(* IEC 61131-3 sources: brOscatLib/oscatBasic (part 6) *)

FUNCTION MIRROR : BOOL (* String *) (* http://www.oscat.de/images/OSCATBasic/oscat_basic333_en.pdf#page=174 *)
	VAR_INPUT
		STR : STRING[STRING_LENGTH];
	END_VAR
	VAR_IN_OUT
		RETVAL : STRING[STRING_LENGTH]; (*Return value of the function*)
	END_VAR
	VAR
		pi : REFERENCE TO ARRAY[1..255] OF BYTE;
		po : REFERENCE TO BYTE;
		lx : INT;
		i : INT;
	END_VAR
END_FUNCTION

FUNCTION MIX : REAL (* Signal processing *) (* http://www.oscat.de/images/OSCATBasic/oscat_basic333_en.pdf#page=281 *)
	VAR_INPUT
		A : REAL;
		B : REAL;
		M : REAL;
	END_VAR
END_FUNCTION

FUNCTION MODR : REAL (* Mathematical *) (* http://www.oscat.de/images/OSCATBasic/oscat_basic333_en.pdf#page=60 *)
	VAR_INPUT
		IN : REAL;
		DIVI : REAL;
	END_VAR
END_FUNCTION

FUNCTION MONTH_BEGIN : DATE (* Time and date *) (* http://www.oscat.de/images/OSCATBasic/oscat_basic333_en.pdf#page=129 *)
	VAR_INPUT
		IDATE : DATE;
	END_VAR
END_FUNCTION

FUNCTION MONTH_END : DATE (* Time and date *) (* http://www.oscat.de/images/OSCATBasic/oscat_basic333_en.pdf#page=130 *)
	VAR_INPUT
		IDATE : DATE;
	END_VAR
END_FUNCTION

FUNCTION MONTH_OF_DATE : INT (* Time and date *) (* http://www.oscat.de/images/OSCATBasic/oscat_basic333_en.pdf#page=130 *)
	VAR_INPUT
		IDATE : DATE;
	END_VAR
END_FUNCTION

FUNCTION MONTH_TO_STRING : BOOL (* String *) (* http://www.oscat.de/images/OSCATBasic/oscat_basic333_en.pdf#page=175 *)
	VAR_INPUT
		MTH : INT;
		LANG : INT;
		LX : INT;
	END_VAR
	VAR_IN_OUT
		RETVAL : STRING[10]; (*Return value of the function*)
	END_VAR
	VAR
		ly : INT;
	END_VAR
	VAR CONSTANT
		cMONTHS : ARRAY[1..3,1..12] OF STRING[10] := ['January','February','March','April','May','June','July','August','September','October','November','December','Januar','Februar','März','April','Mai','Juni','Juli','August','September','Oktober','November','Dezember','Janvier','Février','mars','Avril','Mai','Juin','Juillet','Août','Septembre','Octobre','Novembre','Decembre'];
		cMONTHS3 : ARRAY[1..3,1..12] OF STRING[3] := ['Jan','Feb','Mar','Apr','May','Jun','Jul','Aug','Sep','Oct','Nov','Dec','Jan','Feb','Mrz','Apr','Mai','Jun','Jul','Aug','Sep','Okt','Nov','Dez','Jan','Fev','Mar','Avr','Mai','Jun','Jul','Aou','Sep','Oct','Nov','Dec'];
	END_VAR
END_FUNCTION

FUNCTION MS_TO_BFT : INT (* Conversion *) (* http://www.oscat.de/images/OSCATBasic/oscat_basic333_en.pdf#page=368 *)
	VAR_INPUT
		MS : REAL;
	END_VAR
END_FUNCTION

FUNCTION MS_TO_KMH : REAL (* Conversion *) (* http://www.oscat.de/images/OSCATBasic/oscat_basic333_en.pdf#page=369 *)
	VAR_INPUT
		MS : REAL;
	END_VAR
END_FUNCTION

FUNCTION MULTIME : TIME (* Time and date *) (* http://www.oscat.de/images/OSCATBasic/oscat_basic333_en.pdf#page=130 *)
	VAR_INPUT
		T : TIME;
		M : REAL;
	END_VAR
END_FUNCTION

FUNCTION MULTI_IN : REAL (* Sensor *) (* http://www.oscat.de/images/OSCATBasic/oscat_basic333_en.pdf#page=317 *)
	VAR_INPUT
		IN_1 : REAL;
		IN_2 : REAL;
		IN_3 : REAL;
		DEFAULT : REAL;
		IN_MIN : REAL;
		IN_MAX : REAL;
		MODE : USINT;
	END_VAR
	VAR
		count : INT;
		F1 : BOOL;
		F2 : BOOL;
		F3 : BOOL;
	END_VAR
END_FUNCTION

FUNCTION MUL_ADD : REAL (* Mathematical *) (* http://www.oscat.de/images/OSCATBasic/oscat_basic333_en.pdf#page=61 *)
	VAR_INPUT
		X : REAL;
		K : REAL;
		O : REAL;
	END_VAR
END_FUNCTION

FUNCTION MUX_2 : BOOL (* Gate logic *) (* http://www.oscat.de/images/OSCATBasic/oscat_basic333_en.pdf#page=229 *)
	VAR_INPUT
		D0 : BOOL;
		D1 : BOOL;
		A0 : BOOL;
	END_VAR
END_FUNCTION

FUNCTION MUX_4 : BOOL (* Gate logic *) (* http://www.oscat.de/images/OSCATBasic/oscat_basic333_en.pdf#page=229 *)
	VAR_INPUT
		D0 : BOOL;
		D1 : BOOL;
		D2 : BOOL;
		D3 : BOOL;
		A0 : BOOL;
		A1 : BOOL;
	END_VAR
END_FUNCTION

FUNCTION MUX_R2 : REAL (* Signal processing *) (* http://www.oscat.de/images/OSCATBasic/oscat_basic333_en.pdf#page=281 *)
	VAR_INPUT
		IN0 : REAL;
		IN1 : REAL;
		A : BOOL;
	END_VAR
END_FUNCTION

FUNCTION MUX_R4 : REAL (* Signal processing *) (* http://www.oscat.de/images/OSCATBasic/oscat_basic333_en.pdf#page=282 *)
	VAR_INPUT
		IN0 : REAL;
		IN1 : REAL;
		IN2 : REAL;
		IN3 : REAL;
		A0 : BOOL;
		A1 : BOOL;
	END_VAR
END_FUNCTION

FUNCTION_BLOCK M_D (* Measurements *) (* http://www.oscat.de/images/OSCATBasic/oscat_basic333_en.pdf#page=341 *)
	VAR_INPUT
		START : BOOL;
		STOP : BOOL;
		TMAX : TIME := TIME#14400m0s0ms;
		RST : BOOL;
	END_VAR
	VAR_OUTPUT
		PT : TIME;
		ET : TIME;
		RUN : BOOL;
	END_VAR
	VAR
		edge_ : BOOL;
		T0 : TIME;
		tx : TIME;
		startup : BOOL;
	END_VAR
END_FUNCTION_BLOCK

FUNCTION_BLOCK M_T (* Measurements *) (* http://www.oscat.de/images/OSCATBasic/oscat_basic333_en.pdf#page=342 *)
	VAR_INPUT
		IN : BOOL;
		TMAX : TIME := TIME#14400m0s0ms;
		RST : BOOL;
	END_VAR
	VAR_OUTPUT
		PT : TIME;
		ET : TIME;
	END_VAR
	VAR
		edge_ : BOOL;
		start : TIME;
		tx : TIME;
	END_VAR
END_FUNCTION_BLOCK

FUNCTION_BLOCK M_TX (* Measurements *) (* http://www.oscat.de/images/OSCATBasic/oscat_basic333_en.pdf#page=342 *)
	VAR_INPUT
		IN : BOOL;
		TMAX : TIME := TIME#14400m0s0ms;
		RST : BOOL;
	END_VAR
	VAR_OUTPUT
		TH : TIME;
		TL : TIME;
		DC : REAL;
		F : REAL;
		ET : TIME;
	END_VAR
	VAR
		edge_ : BOOL;
		start : TIME;
		stop : TIME;
		tx : TIME;
		rise : BOOL;
		fall : BOOL;
		startup : BOOL;
	END_VAR
END_FUNCTION_BLOCK

FUNCTION NEGX : REAL (* Mathematical *) (* http://www.oscat.de/images/OSCATBasic/oscat_basic333_en.pdf#page=61 *)
	VAR_INPUT
		X : REAL;
	END_VAR
END_FUNCTION

FUNCTION OCT_TO_BYTE : BYTE (* String *) (* http://www.oscat.de/images/OSCATBasic/oscat_basic333_en.pdf#page=175 *)
	VAR_INPUT
		OCT : STRING[10];
	END_VAR
	VAR
		pt : REFERENCE TO BYTE;
		i : INT;
		X : BYTE;
		stop : INT;
		intX : USINT;
	END_VAR
END_FUNCTION

FUNCTION OCT_TO_DWORD : DWORD (* String *) (* http://www.oscat.de/images/OSCATBasic/oscat_basic333_en.pdf#page=176 *)
	VAR_INPUT
		OCT : STRING[20];
	END_VAR
	VAR
		pt : REFERENCE TO BYTE;
		i : INT;
		X : BYTE;
		stop : INT;
		intX : USINT;
		temp : UDINT;
	END_VAR
END_FUNCTION

FUNCTION OFFSET : REAL (* Signal processing *) (* http://www.oscat.de/images/OSCATBasic/oscat_basic333_en.pdf#page=282 *)
	VAR_INPUT
		X : REAL;
		O1 : BOOL;
		O2 : BOOL;
		O3 : BOOL;
		O4 : BOOL;
		D : BOOL;
		OFFSET_1 : REAL;
		OFFSET_2 : REAL;
		OFFSET_3 : REAL;
		OFFSET_4 : REAL;
		DEFAULT : REAL;
	END_VAR
END_FUNCTION

FUNCTION OFFSET2 : REAL (* Signal processing *) (* http://www.oscat.de/images/OSCATBasic/oscat_basic333_en.pdf#page=285 *)
	VAR_INPUT
		X : REAL;
		O1 : BOOL;
		O2 : BOOL;
		O3 : BOOL;
		O4 : BOOL;
		D : BOOL;
		OFFSET_1 : REAL;
		OFFSET_2 : REAL;
		OFFSET_3 : REAL;
		OFFSET_4 : REAL;
		DEFAULT : REAL;
	END_VAR
END_FUNCTION

FUNCTION OM_TO_F : REAL (* Conversion *) (* http://www.oscat.de/images/OSCATBasic/oscat_basic333_en.pdf#page=369 *)
	VAR_INPUT
		OM : REAL;
	END_VAR
END_FUNCTION

FUNCTION_BLOCK ONTIME (* Measurements *) (* http://www.oscat.de/images/OSCATBasic/oscat_basic333_en.pdf#page=346 *)
	VAR_INPUT
		IN : BOOL;
		RST : BOOL;
	END_VAR
	VAR_IN_OUT
		SECONDS : UDINT;
		CYCLES : UDINT;
	END_VAR
	VAR
		tx : UDINT;
		last : UDINT;
		edge_ : BOOL;
		init : BOOL;
		ms : UDINT;
	END_VAR
END_FUNCTION_BLOCK

FUNCTION OSCAT_VERSION : DWORD (* Other *) (* http://www.oscat.de/images/OSCATBasic/oscat_basic333_en.pdf#page=37 *)
	VAR_INPUT
		IN : BOOL;
	END_VAR
END_FUNCTION

FUNCTION OVERRIDE : REAL (* Signal processing *) (* http://www.oscat.de/images/OSCATBasic/oscat_basic333_en.pdf#page=286 *)
	VAR_INPUT
		X1 : REAL;
		X2 : REAL;
		X3 : REAL;
		E1 : BOOL;
		E2 : BOOL;
		E3 : BOOL;
	END_VAR
END_FUNCTION

FUNCTION PARITY : BOOL (* Gate logic *) (* http://www.oscat.de/images/OSCATBasic/oscat_basic333_en.pdf#page=230 *)
	VAR_INPUT
		IN : DWORD;
	END_VAR
END_FUNCTION

FUNCTION_BLOCK PARSET (* Automation *) (* http://www.oscat.de/images/OSCATBasic/oscat_basic333_en.pdf#page=466 *)
	VAR_INPUT
		A0 : BOOL;
		A1 : BOOL;
		X01 : REAL;
		X02 : REAL;
		X03 : REAL;
		X04 : REAL;
		X11 : REAL;
		X12 : REAL;
		X13 : REAL;
		X14 : REAL;
		X21 : REAL;
		X22 : REAL;
		X23 : REAL;
		X24 : REAL;
		X31 : REAL;
		X32 : REAL;
		X33 : REAL;
		X34 : REAL;
		TC : TIME;
	END_VAR
	VAR_OUTPUT
		P1 : REAL;
		P2 : REAL;
		P3 : REAL;
		P4 : REAL;
	END_VAR
	VAR
		X : ARRAY[0..3,1..4] OF REAL;
		S1 : REAL;
		S2 : REAL;
		S3 : REAL;
		S4 : REAL;
		tx : UDINT;
		last : UDINT;
		start : BOOL;
		set : USINT;
		init : BOOL;
	END_VAR
END_FUNCTION_BLOCK

FUNCTION_BLOCK PARSET2 (* Automation *) (* http://www.oscat.de/images/OSCATBasic/oscat_basic333_en.pdf#page=467 *)
	VAR_INPUT
		X : REAL;
		X01 : REAL;
		X02 : REAL;
		X03 : REAL;
		X04 : REAL;
		X11 : REAL;
		X12 : REAL;
		X13 : REAL;
		X14 : REAL;
		X21 : REAL;
		X22 : REAL;
		X23 : REAL;
		X24 : REAL;
		X31 : REAL;
		X32 : REAL;
		X33 : REAL;
		X34 : REAL;
		L1 : REAL;
		L2 : REAL;
		L3 : REAL;
		TC : TIME;
	END_VAR
	VAR_OUTPUT
		P1 : REAL;
		P2 : REAL;
		P3 : REAL;
		P4 : REAL;
	END_VAR
	VAR
		Pset : PARSET;
		init : BOOL;
	END_VAR
END_FUNCTION_BLOCK

FUNCTION PERIOD : BOOL (* Time and date *) (* http://www.oscat.de/images/OSCATBasic/oscat_basic333_en.pdf#page=131 *)
	VAR_INPUT
		D1 : DATE;
		DX : DATE;
		D2 : DATE;
	END_VAR
	VAR
		day1 : INT;
		day2 : INT;
		dayx : INT;
	END_VAR
END_FUNCTION

FUNCTION PERIOD2 : BOOL (* Time and date *) (* http://www.oscat.de/images/OSCATBasic/oscat_basic333_en.pdf#page=131 *)
	VAR_INPUT
		DP : ARRAY[0..3,0..1] OF DATE;
		DX : DATE;
	END_VAR
END_FUNCTION

FUNCTION_BLOCK PIN_CODE (* Others *) (* http://www.oscat.de/images/OSCATBasic/oscat_basic333_en.pdf#page=231 *)
	VAR_INPUT
		CB : BYTE;
		E : BOOL;
		PIN : STRING[8];
	END_VAR
	VAR_OUTPUT
		TP : BOOL;
	END_VAR
	VAR
		POS : INT := 1;
	END_VAR
END_FUNCTION_BLOCK

FUNCTION POLYNOM_INT : REAL (* Functions *) (* http://www.oscat.de/images/OSCATBasic/oscat_basic333_en.pdf#page=102 *)
	VAR_INPUT
		X : REAL;
		XY : ARRAY[1..5,0..1] OF REAL;
		PTS : INT;
	END_VAR
	VAR
		I : INT;
		J : INT;
		stop : INT;
	END_VAR
END_FUNCTION

FUNCTION_BLOCK PRESSURE (* Conversion *) (* http://www.oscat.de/images/OSCATBasic/oscat_basic333_en.pdf#page=371 *)
	VAR_INPUT
		MWS : REAL;
		TORR : REAL;
		ATT : REAL;
		ATM : REAL;
		PA : REAL;
		BAR : REAL;
	END_VAR
	VAR_OUTPUT
		YMWS : REAL;
		YTORR : REAL;
		YATT : REAL;
		YATM : REAL;
		YPA : REAL;
		YBAR : REAL;
	END_VAR
END_FUNCTION_BLOCK

FUNCTION PT_TO_F : REAL (* Conversion *) (* http://www.oscat.de/images/OSCATBasic/oscat_basic333_en.pdf#page=372 *)
	VAR_INPUT
		PT : TIME;
	END_VAR
END_FUNCTION

FUNCTION_BLOCK PWM_DC (* Signal generators *) (* http://www.oscat.de/images/OSCATBasic/oscat_basic333_en.pdf#page=263 *)
	VAR_INPUT
		F : REAL;
		DC : REAL;
	END_VAR
	VAR_OUTPUT
		Q : BOOL;
	END_VAR
	VAR
		clk : CLK_PRG;
		pulse : TP_X;
		tmp : REAL;
	END_VAR
END_FUNCTION_BLOCK

FUNCTION_BLOCK PWM_PW (* Signal generators *) (* http://www.oscat.de/images/OSCATBasic/oscat_basic333_en.pdf#page=264 *)
	VAR_INPUT
		F : REAL;
		PW : TIME;
	END_VAR
	VAR_OUTPUT
		Q : BOOL;
	END_VAR
	VAR
		clk : CLK_PRG;
		pulse : TP_X;
	END_VAR
END_FUNCTION_BLOCK

FUNCTION R2_ABS : BOOL (* Double Precision *) (* http://www.oscat.de/images/OSCATBasic/oscat_basic333_en.pdf#page=93 *)
	VAR_INPUT
		X : REAL2;
	END_VAR
	VAR_IN_OUT
		RETVAL : REAL2; (*Return value of the function*)
	END_VAR
END_FUNCTION

FUNCTION R2_ADD : BOOL (* Double Precision *) (* http://www.oscat.de/images/OSCATBasic/oscat_basic333_en.pdf#page=93 *)
	VAR_INPUT
		X : REAL2;
		Y : REAL;
	END_VAR
	VAR_IN_OUT
		RETVAL : REAL2; (*Return value of the function*)
	END_VAR
	VAR
		temp : REAL;
	END_VAR
END_FUNCTION

FUNCTION R2_ADD2 : BOOL (* Double Precision *) (* http://www.oscat.de/images/OSCATBasic/oscat_basic333_en.pdf#page=94 *)
	VAR_INPUT
		X : REAL2;
		Y : REAL2;
	END_VAR
	VAR_IN_OUT
		RETVAL : REAL2; (*Return value of the function*)
	END_VAR
END_FUNCTION

FUNCTION R2_MUL : BOOL (* Double Precision *) (* http://www.oscat.de/images/OSCATBasic/oscat_basic333_en.pdf#page=94 *)
	VAR_INPUT
		X : REAL2;
		Y : REAL;
	END_VAR
	VAR_IN_OUT
		RETVAL : REAL2; (*Return value of the function*)
	END_VAR
END_FUNCTION

FUNCTION R2_SET : BOOL (* Double Precision *) (* http://www.oscat.de/images/OSCATBasic/oscat_basic333_en.pdf#page=95 *)
	VAR_INPUT
		X : REAL;
	END_VAR
	VAR_IN_OUT
		RETVAL : REAL2; (*Return value of the function*)
	END_VAR
END_FUNCTION

FUNCTION RAD : REAL (* Mathematical *) (* http://www.oscat.de/images/OSCATBasic/oscat_basic333_en.pdf#page=61 *)
	VAR_INPUT
		DEG : REAL;
	END_VAR
END_FUNCTION

FUNCTION RANGE_TO_BYTE : BYTE (* Signal processing *) (* http://www.oscat.de/images/OSCATBasic/oscat_basic333_en.pdf#page=288 *)
	VAR_INPUT
		X : REAL;
		LOW : REAL;
		HIGH : REAL;
	END_VAR
END_FUNCTION

FUNCTION RANGE_TO_WORD : WORD (* Signal processing *) (* http://www.oscat.de/images/OSCATBasic/oscat_basic333_en.pdf#page=288 *)
	VAR_INPUT
		X : REAL;
		LOW : REAL;
		HIGH : REAL;
	END_VAR
END_FUNCTION

FUNCTION RDM : REAL (* Mathematical *) (* http://www.oscat.de/images/OSCATBasic/oscat_basic333_en.pdf#page=62 *)
	VAR_INPUT
		LAST : REAL;
	END_VAR
	VAR
		tn : UDINT;
		tc : INT;
	END_VAR
END_FUNCTION

FUNCTION RDM2 : INT (* Mathematical *) (* http://www.oscat.de/images/OSCATBasic/oscat_basic333_en.pdf#page=62 *)
	VAR_INPUT
		LAST : INT;
		LOW : INT;
		HIGH : INT;
	END_VAR
END_FUNCTION

FUNCTION RDMDW : DWORD (* Mathematical *) (* http://www.oscat.de/images/OSCATBasic/oscat_basic333_en.pdf#page=63 *)
	VAR_INPUT
		LAST : DWORD;
	END_VAR
	VAR
		RX : REAL;
		M : REAL;
	END_VAR
END_FUNCTION

FUNCTION REAL_TO_DW : DWORD (* Gate logic *) (* http://www.oscat.de/images/OSCATBasic/oscat_basic333_en.pdf#page=231 *)
	VAR_INPUT
		X : REAL;
	END_VAR
	VAR
		pt : REFERENCE TO DWORD;
	END_VAR
END_FUNCTION

FUNCTION REAL_TO_FRAC : BOOL (* Mathematical *) (* http://www.oscat.de/images/OSCATBasic/oscat_basic333_en.pdf#page=64 *)
	VAR_INPUT
		X : REAL; (* in einen Bruch umzuwandelnder Wert *)
		N : INT; (* maximale Größe des Nenners *)
	END_VAR
	VAR_IN_OUT
		RETVAL : FRACTION; (*Return value of the function*)
	END_VAR
	VAR
		temp : DINT; (* Merker für Berechnungen *)
		sign : BOOL; (* Vorzeichen vom Eingangswert *)
		X_gerundet : DINT; (* Wert von Bruch, auf ganze Zahl gerundet *)
		X_ohne_Nachkomma : REAL; (* Wert von Bruch, ohne Nachkommastellen *)
		Numerator : DINT := 1; (* Initialwert Zaehler  *)
		Denominator : DINT := 0; (* Initialwert Nenner *)
		Numerator_old : DINT := 0; (* Initialwert Zaehler der letzten Berechnung  *)
		Denominator_old : DINT := 1; (* Initialwert Zaehler der letzten Berechnung   *)
	END_VAR
END_FUNCTION

FUNCTION REAL_TO_STRF : BOOL (* String *) (* http://www.oscat.de/images/OSCATBasic/oscat_basic333_en.pdf#page=176 *)
	VAR_INPUT
		IN : REAL;
		N : INT;
		D : STRING[1];
	END_VAR
	VAR_IN_OUT
		RETVAL : STRING[20]; (*Return value of the function*)
	END_VAR
	VAR
		O : REAL;
		i : INT;
	END_VAR
END_FUNCTION

FUNCTION REFLECT : DWORD (* Gate logic *) (* http://www.oscat.de/images/OSCATBasic/oscat_basic333_en.pdf#page=232 *)
	VAR_INPUT
		D : DWORD;
		L : INT;
	END_VAR
	VAR
		i : INT;
	END_VAR
END_FUNCTION

FUNCTION REFRACTION : REAL (* Time and date *) (* http://www.oscat.de/images/OSCATBasic/oscat_basic333_en.pdf#page=132 *)
	VAR_INPUT
		ELEV : REAL;
	END_VAR
END_FUNCTION

FUNCTION REPLACE_ALL : BOOL (* String *) (* http://www.oscat.de/images/OSCATBasic/oscat_basic333_en.pdf#page=177 *)
	VAR_INPUT
		STR : STRING[STRING_LENGTH];
		SRC : STRING[STRING_LENGTH];
		REP : STRING[STRING_LENGTH];
	END_VAR
	VAR_IN_OUT
		RETVAL : STRING[STRING_LENGTH]; (*Return value of the function*)
	END_VAR
	VAR
		pos : INT;
		lp : INT;
		lx : INT;
	END_VAR
END_FUNCTION

FUNCTION REPLACE_CHARS : BOOL (* String *) (* http://www.oscat.de/images/OSCATBasic/oscat_basic333_en.pdf#page=177 *)
	VAR_INPUT
		STR : STRING[STRING_LENGTH];
		SRC : STRING[255];
		REP : STRING[255];
	END_VAR
	VAR_IN_OUT
		RETVAL : STRING[STRING_LENGTH]; (*Return value of the function*)
	END_VAR
	VAR
		a : INT;
		b : INT;
		c : STRING[1];
		stp : INT;
	END_VAR
END_FUNCTION

FUNCTION REPLACE_UML : BOOL (* String *) (* http://www.oscat.de/images/OSCATBasic/oscat_basic333_en.pdf#page=178 *)
	VAR_INPUT
		STR : STRING[STRING_LENGTH];
	END_VAR
	VAR_IN_OUT
		RETVAL : STRING[STRING_LENGTH]; (*Return value of the function*)
	END_VAR
	VAR
		L : INT;
		pt : REFERENCE TO BYTE;
		pto : REFERENCE TO BYTE;
		ptm : REFERENCE TO BYTE;
		pt1 : REFERENCE TO BYTE;
		pt2 : REFERENCE TO BYTE;
		su : STRING[2];
		pos : INT;
	END_VAR
END_FUNCTION

FUNCTION RES_NI : REAL (* Sensor *) (* http://www.oscat.de/images/OSCATBasic/oscat_basic333_en.pdf#page=318 *)
	VAR_INPUT
		T : REAL;
		R0 : REAL;
	END_VAR
	VAR CONSTANT
		A : REAL := 0.5485;
		B : REAL := 0.000665;
		C : REAL := 2.805E-09;
	END_VAR
	VAR
		T2 : REAL;
	END_VAR
END_FUNCTION

FUNCTION RES_NTC : REAL (* Sensor *) (* http://www.oscat.de/images/OSCATBasic/oscat_basic333_en.pdf#page=319 *)
	VAR_INPUT
		T : REAL;
		RN : REAL;
		B : REAL;
	END_VAR
END_FUNCTION

FUNCTION RES_PT : REAL (* Sensor *) (* http://www.oscat.de/images/OSCATBasic/oscat_basic333_en.pdf#page=322 *)
	VAR_INPUT
		T : REAL;
		R0 : REAL;
	END_VAR
	VAR CONSTANT
		A : REAL := 0.00390802;
		B : REAL := -5.802E-07;
		C : REAL := -4.2735E-12;
	END_VAR
	VAR
		T2 : REAL;
	END_VAR
END_FUNCTION

FUNCTION RES_SI : REAL (* Sensor *) (* http://www.oscat.de/images/OSCATBasic/oscat_basic333_en.pdf#page=323 *)
	VAR_INPUT
		T : REAL;
		RS : REAL;
		TS : REAL;
	END_VAR
	VAR CONSTANT
		A : REAL := 0.00764;
		B : REAL := 1.66E-05;
	END_VAR
	VAR
		TX : REAL;
	END_VAR
END_FUNCTION

FUNCTION REVERSE : BYTE (* Gate logic *) (* http://www.oscat.de/images/OSCATBasic/oscat_basic333_en.pdf#page=232 *)
	VAR_INPUT
		IN : BYTE;
	END_VAR
END_FUNCTION

FUNCTION_BLOCK RMP_B (* Signal generators *) (* http://www.oscat.de/images/OSCATBasic/oscat_basic333_en.pdf#page=264 *)
	VAR_INPUT
		SET : BOOL;
		PT : TIME;
		E : BOOL := TRUE;
		UP : BOOL := TRUE;
		RST : BOOL;
	END_VAR
	VAR_OUTPUT
		OUT : BYTE;
		BUSY : BOOL;
		HIGH : BOOL;
		LOW : BOOL;
	END_VAR
	VAR
		rmp : _RMP_B;
	END_VAR
END_FUNCTION_BLOCK

FUNCTION_BLOCK RMP_SOFT (* Signal generators *) (* http://www.oscat.de/images/OSCATBasic/oscat_basic333_en.pdf#page=266 *)
	VAR_INPUT
		IN : BOOL;
		VAL : BYTE;
		PT_ON : TIME;
		PT_OFF : TIME;
	END_VAR
	VAR_OUTPUT
		OUT : BYTE;
	END_VAR
	VAR
		rmp : _RMP_B;
		tmp : BYTE;
	END_VAR
END_FUNCTION_BLOCK

FUNCTION_BLOCK RMP_W (* Signal generators *) (* http://www.oscat.de/images/OSCATBasic/oscat_basic333_en.pdf#page=267 *)
	VAR_INPUT
		SET : BOOL;
		PT : TIME;
		E : BOOL := TRUE;
		UP : BOOL := TRUE;
		RST : BOOL;
	END_VAR
	VAR_OUTPUT
		OUT : WORD;
		BUSY : BOOL;
		HIGH : BOOL;
		LOW : BOOL;
	END_VAR
	VAR
		rmp : _RMP_W;
	END_VAR
END_FUNCTION_BLOCK

FUNCTION RND : REAL (* Mathematical *) (* http://www.oscat.de/images/OSCATBasic/oscat_basic333_en.pdf#page=64 *)
	VAR_INPUT
		X : REAL;
		N : INT;
	END_VAR
	VAR
		M : REAL;
	END_VAR
END_FUNCTION

FUNCTION ROUND : REAL (* Mathematical *) (* http://www.oscat.de/images/OSCATBasic/oscat_basic333_en.pdf#page=65 *)
	VAR_INPUT
		IN : REAL;
		N : INT;
	END_VAR
	VAR
		X : REAL;
	END_VAR
	VAR CONSTANT
		cDECADES : ARRAY[0..8] OF REAL := [1,10,100,1000,10000,100000,1000000,10000000,100000000];
	END_VAR
END_FUNCTION

FUNCTION_BLOCK RTC_2 (* Time and date *) (* http://www.oscat.de/images/OSCATBasic/oscat_basic333_en.pdf#page=133 *)
	VAR_INPUT
		SET : BOOL;
		SDT : DATE_AND_TIME;
		SMS : INT;
		DEN : BOOL;
		OFS : INT;
	END_VAR
	VAR_OUTPUT
		UDT : DATE_AND_TIME;
		LOCAL_DT : DATE_AND_TIME;
		DSO : BOOL;
		XMS : INT;
	END_VAR
	VAR
		RT : RTC_MS;
	END_VAR
END_FUNCTION_BLOCK

FUNCTION_BLOCK RTC_MS (* Time and date *) (* http://www.oscat.de/images/OSCATBasic/oscat_basic333_en.pdf#page=134 *)
	VAR_INPUT
		SET : BOOL;
		SDT : DATE_AND_TIME;
		SMS : INT;
	END_VAR
	VAR_OUTPUT
		XDT : DATE_AND_TIME;
		XMS : INT;
	END_VAR
	VAR
		init : BOOL;
		last : UDINT;
		Tx : UDINT;
	END_VAR
END_FUNCTION_BLOCK

FUNCTION SCALE : REAL (* Signal processing *) (* http://www.oscat.de/images/OSCATBasic/oscat_basic333_en.pdf#page=288 *)
	VAR_INPUT
		X : REAL;
		K : REAL;
		O : REAL;
		MX : REAL;
		MN : REAL;
	END_VAR
END_FUNCTION

FUNCTION SCALE_B : REAL (* Signal processing *) (* http://www.oscat.de/images/OSCATBasic/oscat_basic333_en.pdf#page=289 *)
	VAR_INPUT
		X : BYTE;
		I_LO : BYTE;
		I_HI : BYTE;
		O_LO : REAL;
		O_HI : REAL;
	END_VAR
	VAR
		_I_HI : USINT;
		_I_LO : USINT;
	END_VAR
END_FUNCTION

FUNCTION SCALE_B2 : REAL (* Signal processing *) (* http://www.oscat.de/images/OSCATBasic/oscat_basic333_en.pdf#page=290 *)
	VAR_INPUT
		IN1 : BYTE;
		IN2 : BYTE;
		K : REAL;
		O : REAL;
		IN1_MIN : REAL;
		IN1_MAX : REAL := 1000;
		IN2_MIN : REAL;
		IN2_MAX : REAL := 1000;
	END_VAR
END_FUNCTION

FUNCTION SCALE_B4 : REAL (* Signal processing *) (* http://www.oscat.de/images/OSCATBasic/oscat_basic333_en.pdf#page=291 *)
	VAR_INPUT
		IN1 : BYTE;
		IN2 : BYTE;
		IN3 : BYTE;
		IN4 : BYTE;
		K : REAL;
		O : REAL;
		IN1_MIN : REAL;
		IN1_MAX : REAL := 1000;
		IN2_MIN : REAL;
		IN2_MAX : REAL := 1000;
		IN3_MIN : REAL;
		IN3_MAX : REAL := 1000;
		IN4_MIN : REAL;
		IN4_MAX : REAL := 1000;
	END_VAR
END_FUNCTION

FUNCTION SCALE_B8 : REAL (* Signal processing *) (* http://www.oscat.de/images/OSCATBasic/oscat_basic333_en.pdf#page=292 *)
	VAR_INPUT
		IN1 : BYTE;
		IN2 : BYTE;
		IN3 : BYTE;
		IN4 : BYTE;
		IN5 : BYTE;
		IN6 : BYTE;
		IN7 : BYTE;
		IN8 : BYTE;
		K : REAL;
		O : REAL;
		IN1_MIN : REAL;
		IN1_MAX : REAL := 1000;
		IN2_MIN : REAL;
		IN2_MAX : REAL := 1000;
		IN3_MIN : REAL;
		IN3_MAX : REAL := 1000;
		IN4_MIN : REAL;
		IN4_MAX : REAL := 1000;
		IN5_MIN : REAL;
		IN5_MAX : REAL := 1000;
		IN6_MIN : REAL;
		IN6_MAX : REAL := 1000;
		IN7_MIN : REAL;
		IN7_MAX : REAL := 1000;
		IN8_MIN : REAL;
		IN8_MAX : REAL := 1000;
	END_VAR
END_FUNCTION

FUNCTION SCALE_D : REAL (* Signal processing *) (* http://www.oscat.de/images/OSCATBasic/oscat_basic333_en.pdf#page=293 *)
	VAR_INPUT
		X : DWORD;
		I_LO : DWORD;
		I_HI : DWORD;
		O_LO : REAL;
		O_HI : REAL;
	END_VAR
	VAR
		_I_HI : UDINT;
		_I_LO : UDINT;
	END_VAR
END_FUNCTION

FUNCTION SCALE_R : REAL (* Signal processing *) (* http://www.oscat.de/images/OSCATBasic/oscat_basic333_en.pdf#page=294 *)
	VAR_INPUT
		X : REAL;
		I_LO : REAL;
		I_HI : REAL;
		O_LO : REAL;
		O_HI : REAL;
	END_VAR
END_FUNCTION

FUNCTION SCALE_X2 : REAL (* Signal processing *) (* http://www.oscat.de/images/OSCATBasic/oscat_basic333_en.pdf#page=295 *)
	VAR_INPUT
		IN1 : BOOL;
		IN2 : BOOL;
		K : REAL;
		O : REAL;
		IN1_MIN : REAL;
		IN1_MAX : REAL := 1000;
		IN2_MIN : REAL;
		IN2_MAX : REAL := 1000;
	END_VAR
END_FUNCTION

FUNCTION SCALE_X4 : REAL (* Signal processing *) (* http://www.oscat.de/images/OSCATBasic/oscat_basic333_en.pdf#page=296 *)
	VAR_INPUT
		IN1 : BOOL;
		IN2 : BOOL;
		IN3 : BOOL;
		IN4 : BOOL;
		K : REAL;
		O : REAL;
		IN1_MIN : REAL;
		IN1_MAX : REAL := 1000;
		IN2_MIN : REAL;
		IN2_MAX : REAL := 1000;
		IN3_MIN : REAL;
		IN3_MAX : REAL := 1000;
		IN4_MIN : REAL;
		IN4_MAX : REAL := 1000;
	END_VAR
END_FUNCTION

FUNCTION SCALE_X8 : REAL (* Signal processing *) (* http://www.oscat.de/images/OSCATBasic/oscat_basic333_en.pdf#page=297 *)
	VAR_INPUT
		IN1 : BOOL;
		IN2 : BOOL;
		IN3 : BOOL;
		IN4 : BOOL;
		IN5 : BOOL;
		IN6 : BOOL;
		IN7 : BOOL;
		IN8 : BOOL;
		K : REAL;
		O : REAL;
		IN1_MIN : REAL;
		IN1_MAX : REAL := 1000;
		IN2_MIN : REAL;
		IN2_MAX : REAL := 1000;
		IN3_MIN : REAL;
		IN3_MAX : REAL := 1000;
		IN4_MIN : REAL;
		IN4_MAX : REAL := 1000;
		IN5_MIN : REAL;
		IN5_MAX : REAL := 1000;
		IN6_MIN : REAL;
		IN6_MAX : REAL := 1000;
		IN7_MIN : REAL;
		IN7_MAX : REAL := 1000;
		IN8_MIN : REAL;
		IN8_MAX : REAL := 1000;
	END_VAR
END_FUNCTION

FUNCTION_BLOCK SCHEDULER (* Generators *) (* http://www.oscat.de/images/OSCATBasic/oscat_basic333_en.pdf#page=198 *)
	VAR_INPUT
		E0 : BOOL;
		E1 : BOOL;
		E2 : BOOL;
		E3 : BOOL;
		T0 : TIME;
		T1 : TIME;
		T2 : TIME;
		T3 : TIME;
	END_VAR
	VAR_OUTPUT
		Q0 : BOOL;
		Q1 : BOOL;
		Q2 : BOOL;
		Q3 : BOOL;
	END_VAR
	VAR
		init : BOOL;
		s0 : TIME;
		s1 : TIME;
		s2 : TIME;
		s3 : TIME;
		tx : TIME;
		c : INT;
	END_VAR
END_FUNCTION_BLOCK

FUNCTION_BLOCK SCHEDULER_2 (* Generators *) (* http://www.oscat.de/images/OSCATBasic/oscat_basic333_en.pdf#page=198 *)
	VAR_INPUT
		E0 : BOOL;
		E1 : BOOL;
		E2 : BOOL;
		E3 : BOOL;
		C0 : UINT;
		C1 : UINT;
		C2 : UINT;
		C3 : UINT;
		O0 : UINT;
		O1 : UINT;
		O2 : UINT;
		O3 : UINT;
	END_VAR
	VAR_OUTPUT
		Q0 : BOOL;
		Q1 : BOOL;
		Q2 : BOOL;
		Q3 : BOOL;
	END_VAR
	VAR
		sx : UINT;
	END_VAR
END_FUNCTION_BLOCK

FUNCTION SDT_TO_DATE : DATE (* Time and date *) (* http://www.oscat.de/images/OSCATBasic/oscat_basic333_en.pdf#page=134 *)
	VAR_INPUT
		DTI : SDT;
	END_VAR
END_FUNCTION

FUNCTION SDT_TO_DT : DATE_AND_TIME (* Time and date *) (* http://www.oscat.de/images/OSCATBasic/oscat_basic333_en.pdf#page=135 *)
	VAR_INPUT
		DTI : SDT;
	END_VAR
END_FUNCTION

FUNCTION SDT_TO_TOD : TIME_OF_DAY (* Time and date *) (* http://www.oscat.de/images/OSCATBasic/oscat_basic333_en.pdf#page=135 *)
	VAR_INPUT
		DTI : SDT;
	END_VAR
END_FUNCTION

FUNCTION SECOND : REAL (* Time and date *) (* http://www.oscat.de/images/OSCATBasic/oscat_basic333_en.pdf#page=135 *)
	VAR_INPUT
		ITOD : TIME_OF_DAY;
	END_VAR
END_FUNCTION

FUNCTION SECOND_OF_DT : INT (* Time and date *) (* http://www.oscat.de/images/OSCATBasic/oscat_basic333_en.pdf#page=136 *)
	VAR_INPUT
		XDT : DATE_AND_TIME;
	END_VAR
END_FUNCTION

FUNCTION SECOND_TO_TIME : TIME (* Time and date *) (* http://www.oscat.de/images/OSCATBasic/oscat_basic333_en.pdf#page=136 *)
	VAR_INPUT
		IN : REAL;
	END_VAR
END_FUNCTION

FUNCTION_BLOCK SEL2_OF_3 (* Signal processing *) (* http://www.oscat.de/images/OSCATBasic/oscat_basic333_en.pdf#page=298 *)
	VAR_INPUT
		IN1 : REAL;
		IN2 : REAL;
		IN3 : REAL;
		D : REAL;
	END_VAR
	VAR_OUTPUT
		Y : REAL;
		W : INT;
		E : BOOL;
	END_VAR
	VAR
		D12 : BOOL;
		D23 : BOOL;
		D31 : BOOL;
	END_VAR
END_FUNCTION_BLOCK

FUNCTION_BLOCK SEL2_OF_3B (* Signal processing *) (* http://www.oscat.de/images/OSCATBasic/oscat_basic333_en.pdf#page=299 *)
	VAR_INPUT
		IN1 : BOOL;
		IN2 : BOOL;
		IN3 : BOOL;
		TD : TIME;
	END_VAR
	VAR_OUTPUT
		Q : BOOL;
		W : BOOL;
	END_VAR
	VAR
		TDEL : TON;
	END_VAR
END_FUNCTION_BLOCK

FUNCTION_BLOCK SELECT_8 (* FF Edge triggered *) (* http://www.oscat.de/images/OSCATBasic/oscat_basic333_en.pdf#page=247 *)
	VAR_INPUT
		E : BOOL;
		SET : BOOL;
		IN : BYTE;
		UP : BOOL;
		DN : BOOL;
		RST : BOOL;
	END_VAR
	VAR_OUTPUT
		Q0 : BOOL;
		Q1 : BOOL;
		Q2 : BOOL;
		Q3 : BOOL;
		Q4 : BOOL;
		Q5 : BOOL;
		Q6 : BOOL;
		Q7 : BOOL;
		STATE : INT;
	END_VAR
	VAR
		last_up : BOOL;
		last_dn : BOOL;
	END_VAR
END_FUNCTION_BLOCK

FUNCTION SENSOR_INT : REAL (* Sensor *) (* http://www.oscat.de/images/OSCATBasic/oscat_basic333_en.pdf#page=324 *)
	VAR_INPUT
		VOLTAGE : REAL;
		CURRENT : REAL;
		RP : REAL;
		RS : REAL;
	END_VAR
	VAR
		RG : REAL;
	END_VAR
END_FUNCTION

FUNCTION_BLOCK SEQUENCE_4 (* Generators *) (* http://www.oscat.de/images/OSCATBasic/oscat_basic333_en.pdf#page=199 *)
	VAR_INPUT
		IN0 : BOOL := TRUE;
		IN1 : BOOL := TRUE;
		IN2 : BOOL := TRUE;
		IN3 : BOOL := TRUE;
		START : BOOL;
		RST : BOOL;
		WAIT0 : TIME;
		DELAY0 : TIME;
		WAIT1 : TIME;
		DELAY1 : TIME;
		WAIT2 : TIME;
		DELAY2 : TIME;
		WAIT3 : TIME;
		DELAY3 : TIME;
		STOP_ON_ERROR : BOOL;
	END_VAR
	VAR_OUTPUT
		Q0 : BOOL;
		Q1 : BOOL;
		Q2 : BOOL;
		Q3 : BOOL;
		QX : BOOL;
		RUN : BOOL;
		STEP : INT := -1;
		STATUS : BYTE;
	END_VAR
	VAR
		last : TIME;
		edge_ : BOOL;
		tx : TIME;
		init : BOOL;
	END_VAR
END_FUNCTION_BLOCK

FUNCTION_BLOCK SEQUENCE_8 (* Generators *) (* http://www.oscat.de/images/OSCATBasic/oscat_basic333_en.pdf#page=203 *)
	VAR_INPUT
		IN0 : BOOL := TRUE;
		IN1 : BOOL := TRUE;
		IN2 : BOOL := TRUE;
		IN3 : BOOL := TRUE;
		IN4 : BOOL := TRUE;
		IN5 : BOOL := TRUE;
		IN6 : BOOL := TRUE;
		IN7 : BOOL := TRUE;
		START : BOOL;
		RST : BOOL;
		WAIT0 : TIME;
		DELAY0 : TIME;
		WAIT1 : TIME;
		DELAY1 : TIME;
		WAIT2 : TIME;
		DELAY2 : TIME;
		WAIT3 : TIME;
		DELAY3 : TIME;
		WAIT4 : TIME;
		DELAY4 : TIME;
		WAIT5 : TIME;
		DELAY5 : TIME;
		WAIT6 : TIME;
		DELAY6 : TIME;
		WAIT7 : TIME;
		DELAY7 : TIME;
		STOP_ON_ERROR : BOOL;
	END_VAR
	VAR_OUTPUT
		Q0 : BOOL;
		Q1 : BOOL;
		Q2 : BOOL;
		Q3 : BOOL;
		Q4 : BOOL;
		Q5 : BOOL;
		Q6 : BOOL;
		Q7 : BOOL;
		QX : BOOL;
		RUN : BOOL;
		STEP : INT := -1;
		STATUS : BYTE;
	END_VAR
	VAR
		last : TIME;
		edge_ : BOOL;
		tx : TIME;
		init : BOOL;
	END_VAR
END_FUNCTION_BLOCK

FUNCTION_BLOCK SEQUENCE_64 (* Generators *) (* http://www.oscat.de/images/OSCATBasic/oscat_basic333_en.pdf#page=202 *)
	VAR_INPUT
		START : BOOL;
		SMAX : INT;
		PROG : ARRAY[0..63] OF TIME;
		RST : BOOL;
	END_VAR
	VAR_OUTPUT
		STATE : INT := -1;
		TRIG : BOOL;
	END_VAR
	VAR
		tx : TIME;
		edge_ : BOOL;
		last : TIME;
	END_VAR
END_FUNCTION_BLOCK

FUNCTION SET_DATE : DATE (* Time and date *) (* http://www.oscat.de/images/OSCATBasic/oscat_basic333_en.pdf#page=136 *)
	VAR_INPUT
		YEAR : INT;
		MONTH : INT;
		DAY : INT;
	END_VAR
	VAR
		count : INT;
		ofs : ARRAY[1..12] OF INT := [0,31,59,90,120,151,181,212,243,273,304,334];
		ENDIF : BOOL;
	END_VAR
END_FUNCTION

FUNCTION SET_DT : DATE_AND_TIME (* Time and date *) (* http://www.oscat.de/images/OSCATBasic/oscat_basic333_en.pdf#page=137 *)
	VAR_INPUT
		YEAR : INT;
		MONTH : INT;
		DAY : INT;
		HOUR : INT;
		MINUTE : INT;
		SECOND : INT;
	END_VAR
END_FUNCTION

FUNCTION SET_TOD : TIME_OF_DAY (* Time and date *) (* http://www.oscat.de/images/OSCATBasic/oscat_basic333_en.pdf#page=138 *)
	VAR_INPUT
		HOUR : INT;
		MINUTE : INT;
		SECOND : REAL;
	END_VAR
END_FUNCTION

FUNCTION SGN : INT (* Mathematical *) (* http://www.oscat.de/images/OSCATBasic/oscat_basic333_en.pdf#page=65 *)
	VAR_INPUT
		X : REAL;
	END_VAR
END_FUNCTION

FUNCTION_BLOCK SH (* Signal processing *) (* http://www.oscat.de/images/OSCATBasic/oscat_basic333_en.pdf#page=299 *)
	VAR_INPUT
		IN : REAL;
		CLK : BOOL;
	END_VAR
	VAR_OUTPUT
		OUT : REAL;
		TRIG : BOOL;
	END_VAR
	VAR
		edge_ : BOOL;
	END_VAR
END_FUNCTION_BLOCK

FUNCTION SHL1 : DWORD (* Gate logic *) (* http://www.oscat.de/images/OSCATBasic/oscat_basic333_en.pdf#page=233 *)
	VAR_INPUT
		IN : DWORD;
		N : INT;
	END_VAR
	VAR CONSTANT
		temp : DWORD := 16#FFFFFFFF;
	END_VAR
END_FUNCTION

FUNCTION SHR1 : DWORD (* Gate logic *) (* http://www.oscat.de/images/OSCATBasic/oscat_basic333_en.pdf#page=233 *)
	VAR_INPUT
		IN : DWORD;
		N : INT;
	END_VAR
	VAR CONSTANT
		temp : DWORD := 16#FFFFFFFF;
	END_VAR
END_FUNCTION

FUNCTION_BLOCK SHR_4E (* FF Edge triggered *) (* http://www.oscat.de/images/OSCATBasic/oscat_basic333_en.pdf#page=249 *)
	VAR_INPUT
		SET : BOOL;
		D0 : BOOL;
		CLK : BOOL;
		RST : BOOL;
	END_VAR
	VAR_OUTPUT
		Q0 : BOOL;
		Q1 : BOOL;
		Q2 : BOOL;
		Q3 : BOOL;
	END_VAR
	VAR
		trig : R_TRIG;
	END_VAR
END_FUNCTION_BLOCK

FUNCTION_BLOCK SHR_4UDE (* FF Edge triggered *) (* http://www.oscat.de/images/OSCATBasic/oscat_basic333_en.pdf#page=250 *)
	VAR_INPUT
		SET : BOOL;
		D0 : BOOL;
		D3 : BOOL;
		CLK : BOOL;
		DN : BOOL;
		RST : BOOL;
	END_VAR
	VAR_OUTPUT
		Q0 : BOOL;
		Q1 : BOOL;
		Q2 : BOOL;
		Q3 : BOOL;
	END_VAR
	VAR
		trig : R_TRIG;
	END_VAR
END_FUNCTION_BLOCK

FUNCTION_BLOCK SHR_8PLE (* FF Edge triggered *) (* http://www.oscat.de/images/OSCATBasic/oscat_basic333_en.pdf#page=251 *)
	VAR_INPUT
		DIN : BOOL;
		DLOAD : BYTE;
		CLK : BOOL;
		UP : BOOL := 1;
		LOAD : BOOL;
		RST : BOOL;
	END_VAR
	VAR_OUTPUT
		DOUT : BOOL;
	END_VAR
	VAR
		edge_ : BOOL := 1;
		register : BYTE;
	END_VAR
END_FUNCTION_BLOCK

FUNCTION_BLOCK SHR_8UDE (* FF Edge triggered *) (* http://www.oscat.de/images/OSCATBasic/oscat_basic333_en.pdf#page=252 *)
	VAR_INPUT
		SET : BOOL;
		D0 : BOOL;
		D7 : BOOL;
		CLK : BOOL;
		DN : BOOL;
		RST : BOOL;
	END_VAR
	VAR_OUTPUT
		Q0 : BOOL;
		Q1 : BOOL;
		Q2 : BOOL;
		Q3 : BOOL;
		Q4 : BOOL;
		Q5 : BOOL;
		Q6 : BOOL;
		Q7 : BOOL;
	END_VAR
	VAR
		trig : R_TRIG;
	END_VAR
END_FUNCTION_BLOCK

FUNCTION_BLOCK SH_1 (* Signal processing *) (* http://www.oscat.de/images/OSCATBasic/oscat_basic333_en.pdf#page=300 *)
	VAR_INPUT
		IN : REAL;
		PT : TIME;
	END_VAR
	VAR_OUTPUT
		OUT : REAL;
		TRIG : BOOL;
	END_VAR
	VAR
		last : TIME;
		tx : TIME;
	END_VAR
END_FUNCTION_BLOCK

FUNCTION_BLOCK SH_2 (* Signal processing *) (* http://www.oscat.de/images/OSCATBasic/oscat_basic333_en.pdf#page=301 *)
	VAR_INPUT
		IN : REAL;
		PT : TIME;
		N : INT := 16;
		DISC : INT;
	END_VAR
	VAR_OUTPUT
		OUT : REAL;
		TRIG : BOOL;
		AVG : REAL;
		HIGH : REAL;
		LOW : REAL;
	END_VAR
	VAR
		M : INT;
		buf : ARRAY[0..15] OF REAL;
		buf2 : ARRAY[0..15] OF REAL;
		last : TIME;
		i : INT;
		start : INT;
		temp : REAL;
		stop : INT;
		tx : TIME;
		d2 : INT;
	END_VAR
END_FUNCTION_BLOCK

FUNCTION_BLOCK SH_T (* Signal processing *) (* http://www.oscat.de/images/OSCATBasic/oscat_basic333_en.pdf#page=303 *)
	VAR_INPUT
		IN : REAL;
		E : BOOL;
	END_VAR
	VAR_OUTPUT
		OUT : REAL;
	END_VAR
END_FUNCTION_BLOCK

FUNCTION SIGMOID : REAL (* Mathematical *) (* http://www.oscat.de/images/OSCATBasic/oscat_basic333_en.pdf#page=66 *)
	VAR_INPUT
		X : REAL;
	END_VAR
END_FUNCTION

FUNCTION_BLOCK SIGNAL (* Automation *) (* http://www.oscat.de/images/OSCATBasic/oscat_basic333_en.pdf#page=468 *)
	VAR_INPUT
		IN : BOOL;
		SIG : BYTE;
		TS : TIME;
	END_VAR
	VAR_OUTPUT
		Q : BOOL;
	END_VAR
	VAR
		tx : UDINT;
		step : BYTE;
	END_VAR
	VAR CONSTANT
		one : BYTE := 1;
	END_VAR
END_FUNCTION_BLOCK

FUNCTION_BLOCK SIGNAL_4 (* Automation *) (* http://www.oscat.de/images/OSCATBasic/oscat_basic333_en.pdf#page=469 *)
	VAR_INPUT
		IN1 : BOOL;
		IN2 : BOOL;
		IN3 : BOOL;
		IN4 : BOOL;
		TS : TIME;
		S1 : BYTE := 2#11111111;
		S2 : BYTE := 2#11110000;
		S3 : BYTE := 2#10101010;
		S4 : BYTE := 2#10100000;
	END_VAR
	VAR_OUTPUT
		Q : BOOL;
	END_VAR
	VAR
		sig : SIGNAL;
	END_VAR
END_FUNCTION_BLOCK

FUNCTION SIGN_I : BOOL (* Mathematical *) (* http://www.oscat.de/images/OSCATBasic/oscat_basic333_en.pdf#page=66 *)
	VAR_INPUT
		IN : DINT;
	END_VAR
END_FUNCTION

FUNCTION SIGN_R : BOOL (* Mathematical *) (* http://www.oscat.de/images/OSCATBasic/oscat_basic333_en.pdf#page=67 *)
	VAR_INPUT
		IN : REAL;
	END_VAR
END_FUNCTION

FUNCTION SINC : REAL (* Mathematical *) (* http://www.oscat.de/images/OSCATBasic/oscat_basic333_en.pdf#page=67 *)
	VAR_INPUT
		X : REAL;
	END_VAR
END_FUNCTION

FUNCTION SINH : REAL (* Mathematical *) (* http://www.oscat.de/images/OSCATBasic/oscat_basic333_en.pdf#page=67 *)
	VAR_INPUT
		X : REAL;
	END_VAR
END_FUNCTION

FUNCTION_BLOCK SPEED (* Conversion *) (* http://www.oscat.de/images/OSCATBasic/oscat_basic333_en.pdf#page=372 *)
	VAR_INPUT
		MS : REAL;
		KMH : REAL;
		KN : REAL;
		MH : REAL;
	END_VAR
	VAR_OUTPUT
		YMS : REAL;
		YKMH : REAL;
		YKN : REAL;
		YMH : REAL;
	END_VAR
END_FUNCTION_BLOCK

FUNCTION SPHERE_V : REAL (* Geometry *) (* http://www.oscat.de/images/OSCATBasic/oscat_basic333_en.pdf#page=106 *)
	VAR_INPUT
		RX : REAL;
	END_VAR
END_FUNCTION

FUNCTION SQRTN : REAL (* Mathematical *) (* http://www.oscat.de/images/OSCATBasic/oscat_basic333_en.pdf#page=68 *)
	VAR_INPUT
		X : REAL;
		N : INT;
	END_VAR
END_FUNCTION

FUNCTION_BLOCK SRAMP (* Automation *) (* http://www.oscat.de/images/OSCATBasic/oscat_basic333_en.pdf#page=470 *)
	VAR_INPUT
		X : REAL;
		A_UP : REAL;
		A_DN : REAL;
		VU_MAX : REAL;
		VD_MAX : REAL;
		LIMIT_HIGH : REAL;
		LIMIT_LOW : REAL;
		RST : BOOL;
	END_VAR
	VAR_OUTPUT
		Y : REAL;
		V : REAL;
	END_VAR
	VAR
		cycle_time : TC_S;
		init : BOOL;
	END_VAR
END_FUNCTION_BLOCK

FUNCTION_BLOCK STACK_16 (* Memory *) (* http://www.oscat.de/images/OSCATBasic/oscat_basic333_en.pdf#page=185 *)
	VAR_INPUT
		DIN : DWORD;
		E : BOOL := TRUE;
		RD : BOOL;
		WD : BOOL;
		RST : BOOL;
	END_VAR
	VAR_OUTPUT
		DOUT : DWORD;
		EMPTY : BOOL := TRUE;
		FULL : BOOL;
	END_VAR
	VAR
		stack : ARRAY[0..n] OF DWORD;
		pt : INT;
	END_VAR
	VAR CONSTANT
		n : INT := 15; (* changing this value will chage the number of stored elements in the fifo *)
	END_VAR
END_FUNCTION_BLOCK

FUNCTION_BLOCK STACK_32 (* Memory *) (* http://www.oscat.de/images/OSCATBasic/oscat_basic333_en.pdf#page=186 *)
	VAR_INPUT
		DIN : DWORD;
		E : BOOL := TRUE;
		RD : BOOL;
		WD : BOOL;
		RST : BOOL;
	END_VAR
	VAR_OUTPUT
		DOUT : DWORD;
		EMPTY : BOOL := TRUE;
		FULL : BOOL;
	END_VAR
	VAR
		stack : ARRAY[0..n] OF DWORD;
		pt : INT;
	END_VAR
	VAR CONSTANT
		n : INT := 31; (* changing this value will chage the number of stored elements in the fifo *)
	END_VAR
END_FUNCTION_BLOCK

FUNCTION STAIR : REAL (* Signal processing *) (* http://www.oscat.de/images/OSCATBasic/oscat_basic333_en.pdf#page=304 *)
	VAR_INPUT
		X : REAL;
		D : REAL;
	END_VAR
END_FUNCTION

FUNCTION_BLOCK STAIR2 (* Signal processing *) (* http://www.oscat.de/images/OSCATBasic/oscat_basic333_en.pdf#page=304 *)
	VAR_INPUT
		X : REAL;
		D : REAL;
	END_VAR
	VAR_OUTPUT
		Y : REAL;
	END_VAR
END_FUNCTION_BLOCK

FUNCTION STATUS_TO_ESR : BOOL (* Other *) (* http://www.oscat.de/images/OSCATBasic/oscat_basic333_en.pdf#page=38 *)
	VAR_INPUT
		STATUS : BYTE;
		ADRESS : STRING[10];
		DT_IN : DATE_AND_TIME;
		TS : TIME;
	END_VAR
	VAR_IN_OUT
		RETVAL : ESR_DATA; (*Return value of the function*)
	END_VAR
END_FUNCTION

FUNCTION_BLOCK STORE_8 (* FF pulse triggered *) (* http://www.oscat.de/images/OSCATBasic/oscat_basic333_en.pdf#page=253 *)
	VAR_INPUT
		SET : BOOL;
		D0 : BOOL;
		D1 : BOOL;
		D2 : BOOL;
		D3 : BOOL;
		D4 : BOOL;
		D5 : BOOL;
		D6 : BOOL;
		D7 : BOOL;
		CLR : BOOL;
		RST : BOOL;
	END_VAR
	VAR_OUTPUT
		Q0 : BOOL;
		Q1 : BOOL;
		Q2 : BOOL;
		Q3 : BOOL;
		Q4 : BOOL;
		Q5 : BOOL;
		Q6 : BOOL;
		Q7 : BOOL;
	END_VAR
	VAR
		edge_ : BOOL;
	END_VAR
END_FUNCTION_BLOCK

FUNCTION SUN_MIDDAY : TIME_OF_DAY (* Time and date *) (* http://www.oscat.de/images/OSCATBasic/oscat_basic333_en.pdf#page=138 *)
	VAR_INPUT
		LON : REAL;
		UTC : DATE;
	END_VAR
	VAR
		T : REAL;
		OFFSET : REAL;
	END_VAR
END_FUNCTION

FUNCTION_BLOCK SUN_POS (* Time and date *) (* http://www.oscat.de/images/OSCATBasic/oscat_basic333_en.pdf#page=138 *)
	VAR_INPUT
		LATITUDE : REAL; (* latitude of geographical position  *)
		LONGITUDE : REAL; (* longitude of geographical position  *)
		UTC : DATE_AND_TIME; (*	world time				*)
	END_VAR
	VAR_OUTPUT
		B : REAL;
		H : REAL;
		HR : REAL;
	END_VAR
	VAR
		g : REAL;
		a : REAL;
		d : REAL;
		t1 : REAL;
		n : REAL;
		e : REAL;
		c : REAL;
		tau : REAL;
		sin_d : REAL;
		rlat : REAL;
		sin_lat : REAL;
		cos_lat : REAL;
		cos_tau : REAL;
		cos_d : REAL;
	END_VAR
END_FUNCTION_BLOCK

FUNCTION_BLOCK SUN_TIME (* Time and date *) (* http://www.oscat.de/images/OSCATBasic/oscat_basic333_en.pdf#page=139 *)
	VAR_INPUT
		LATITUDE : REAL; (* latitude of geographical position  *)
		LONGITUDE : REAL; (* longitude of geographical position  *)
		UTC : DATE; (*	world time	*)
		H : REAL := -0.83333333333; (* heighth above horizon for sunrise *)
	END_VAR
	VAR_OUTPUT
		MIDDAY : TIME_OF_DAY; (*	astrological midday in hours when sun stands at south direction	*)
		SUN_RISE : TIME_OF_DAY; (*	sun rise for current day in local time *)
		SUN_SET : TIME_OF_DAY; (*	sun set for current day in local time *)
		SUN_DECLINATION : REAL; (*	sun declination above horizon at midday in degrees	*)
	END_VAR
	VAR
		dk : REAL; (* sun declination at midday *)
		delta : TIME; (* delta from midday for sunrise and sunset  *)
		b : REAL;
	END_VAR
END_FUNCTION_BLOCK

FUNCTION SWAP_BYTE : WORD (* Gate logic *) (* http://www.oscat.de/images/OSCATBasic/oscat_basic333_en.pdf#page=234 *)
	VAR_INPUT
		IN : WORD;
	END_VAR
END_FUNCTION

FUNCTION SWAP_BYTE2 : DWORD (* Gate logic *) (* http://www.oscat.de/images/OSCATBasic/oscat_basic333_en.pdf#page=234 *)
	VAR_INPUT
		IN : DWORD;
	END_VAR
END_FUNCTION

FUNCTION TANC : REAL (* Mathematical *) (* http://www.oscat.de/images/OSCATBasic/oscat_basic333_en.pdf#page=68 *)
	VAR_INPUT
		X : REAL;
	END_VAR
END_FUNCTION

FUNCTION TANH : REAL (* Mathematical *) (* http://www.oscat.de/images/OSCATBasic/oscat_basic333_en.pdf#page=69 *)
	VAR_INPUT
		X : REAL;
	END_VAR
END_FUNCTION

FUNCTION_BLOCK TC_MS (* Measurements *) (* http://www.oscat.de/images/OSCATBasic/oscat_basic333_en.pdf#page=352 *)
	VAR_OUTPUT
		TC : UDINT;
	END_VAR
	VAR
		init : BOOL;
		tx : UDINT;
		last : UDINT;
	END_VAR
END_FUNCTION_BLOCK

FUNCTION_BLOCK TC_S (* Measurements *) (* http://www.oscat.de/images/OSCATBasic/oscat_basic333_en.pdf#page=353 *)
	VAR_OUTPUT
		TC : REAL;
	END_VAR
	VAR
		init : BOOL;
		tx : UDINT;
		last : UDINT;
	END_VAR
END_FUNCTION_BLOCK

FUNCTION_BLOCK TC_US (* Measurements *) (* http://www.oscat.de/images/OSCATBasic/oscat_basic333_en.pdf#page=353 *)
	VAR_OUTPUT
		TC : UDINT;
	END_VAR
	VAR
		init : BOOL;
		tx : UDINT;
		last : UDINT;
	END_VAR
END_FUNCTION_BLOCK

FUNCTION_BLOCK TEMPERATURE (* Conversion *) (* http://www.oscat.de/images/OSCATBasic/oscat_basic333_en.pdf#page=374 *)
	VAR_INPUT
		K : REAL;
		C : REAL := -273.15;
		F : REAL := -459.67;
		RE : REAL := -218.52;
		RA : REAL;
	END_VAR
	VAR_OUTPUT
		YK : REAL;
		YC : REAL;
		YF : REAL;
		YRE : REAL;
		YRA : REAL;
	END_VAR
END_FUNCTION_BLOCK

FUNCTION TEMP_NI : REAL (* Sensor *) (* http://www.oscat.de/images/OSCATBasic/oscat_basic333_en.pdf#page=325 *)
	VAR_INPUT
		RES : REAL;
		R0 : REAL;
	END_VAR
END_FUNCTION

FUNCTION TEMP_NTC : REAL (* Sensor *) (* http://www.oscat.de/images/OSCATBasic/oscat_basic333_en.pdf#page=326 *)
	VAR_INPUT
		RES : REAL;
		RN : REAL;
		B : REAL;
	END_VAR
END_FUNCTION

FUNCTION TEMP_PT : REAL (* Sensor *) (* http://www.oscat.de/images/OSCATBasic/oscat_basic333_en.pdf#page=326 *)
	VAR_INPUT
		RES : REAL;
		R0 : REAL;
	END_VAR
	VAR CONSTANT
		A : REAL := 0.0039083;
		B : REAL := -5.775E-07;
		accuracy : REAL := 0.01;
	END_VAR
	VAR
		step : REAL := 50;
		X : REAL;
		Y : REAL;
		t1 : REAL;
		pt : REFERENCE TO UDINT;
	END_VAR
END_FUNCTION

FUNCTION TEMP_SI : REAL (* Sensor *) (* http://www.oscat.de/images/OSCATBasic/oscat_basic333_en.pdf#page=331 *)
	VAR_INPUT
		RES : REAL;
		RS : REAL;
		TS : REAL;
	END_VAR
END_FUNCTION

FUNCTION_BLOCK TICKER (* String *) (* http://www.oscat.de/images/OSCATBasic/oscat_basic333_en.pdf#page=178 *)
	VAR_INPUT
		N : INT;
		PT : TIME;
	END_VAR
	VAR_OUTPUT
		DISPLAY : STRING[STRING_LENGTH];
	END_VAR
	VAR_IN_OUT
		TEXT : STRING[STRING_LENGTH];
	END_VAR
	VAR
		delay : TP;
		step : INT;
	END_VAR
END_FUNCTION_BLOCK

FUNCTION TIMECHECK : BOOL (* Time and date *) (* http://www.oscat.de/images/OSCATBasic/oscat_basic333_en.pdf#page=141 *)
	VAR_INPUT
		TD : TIME_OF_DAY;
		START : TIME_OF_DAY;
		STOP : TIME_OF_DAY;
	END_VAR
END_FUNCTION

FUNCTION_BLOCK TMAX (* Generators *) (* http://www.oscat.de/images/OSCATBasic/oscat_basic333_en.pdf#page=204 *)
	VAR_INPUT
		IN : BOOL;
		PT : TIME;
	END_VAR
	VAR_OUTPUT
		Q : BOOL;
		Z : BOOL;
	END_VAR
	VAR
		tx : TIME;
		start : TIME;
		last_in : BOOL;
	END_VAR
END_FUNCTION_BLOCK

FUNCTION_BLOCK TMIN (* Generators *) (* http://www.oscat.de/images/OSCATBasic/oscat_basic333_en.pdf#page=205 *)
	VAR_INPUT
		IN : BOOL;
		PT : TIME;
	END_VAR
	VAR_OUTPUT
		Q : BOOL;
	END_VAR
	VAR
		pm : TP;
	END_VAR
END_FUNCTION_BLOCK

FUNCTION_BLOCK TOF_1 (* Generators *) (* http://www.oscat.de/images/OSCATBasic/oscat_basic333_en.pdf#page=205 *)
	VAR_INPUT
		IN : BOOL;
		PT : TIME;
		RST : BOOL;
	END_VAR
	VAR_OUTPUT
		Q : BOOL;
	END_VAR
	VAR
		tx : TIME;
		start : TIME;
	END_VAR
END_FUNCTION_BLOCK

FUNCTION_BLOCK TOGGLE (* FF Edge triggered *) (* http://www.oscat.de/images/OSCATBasic/oscat_basic333_en.pdf#page=254 *)
	VAR_INPUT
		CLK : BOOL;
		RST : BOOL;
	END_VAR
	VAR_OUTPUT
		Q : BOOL;
	END_VAR
	VAR
		edge_ : BOOL;
	END_VAR
END_FUNCTION_BLOCK

FUNCTION_BLOCK TONOF (* Generators *) (* http://www.oscat.de/images/OSCATBasic/oscat_basic333_en.pdf#page=206 *)
	VAR_INPUT
		IN : BOOL;
		T_ON : TIME;
		T_OFF : TIME;
	END_VAR
	VAR_OUTPUT
		Q : BOOL;
	END_VAR
	VAR
		X : TON;
		old : BOOL;
		mode : BOOL;
	END_VAR
END_FUNCTION_BLOCK

FUNCTION TO_LOWER : BYTE (* String *) (* http://www.oscat.de/images/OSCATBasic/oscat_basic333_en.pdf#page=179 *)
	VAR_INPUT
		IN : BYTE;
	END_VAR
	VAR
		byteAsInt : USINT;
	END_VAR
END_FUNCTION

FUNCTION TO_UML : BOOL (* String *) (* http://www.oscat.de/images/OSCATBasic/oscat_basic333_en.pdf#page=180 *)
	VAR_INPUT
		IN : BYTE;
	END_VAR
	VAR_IN_OUT
		RETVAL : STRING[2]; (*Return value of the function*)
	END_VAR
END_FUNCTION

FUNCTION TO_UPPER : BYTE (* String *) (* http://www.oscat.de/images/OSCATBasic/oscat_basic333_en.pdf#page=180 *)
	VAR_INPUT
		IN : BYTE;
	END_VAR
	VAR
		byteAsInt : USINT;
	END_VAR
END_FUNCTION

FUNCTION_BLOCK TP_1 (* Generators *) (* http://www.oscat.de/images/OSCATBasic/oscat_basic333_en.pdf#page=207 *)
	VAR_INPUT
		IN : BOOL;
		PT : TIME;
		RST : BOOL;
	END_VAR
	VAR_OUTPUT
		Q : BOOL;
	END_VAR
	VAR
		tx : TIME;
		start : TIME;
		ix : BOOL;
	END_VAR
END_FUNCTION_BLOCK

FUNCTION_BLOCK TP_1D (* Generators *) (* http://www.oscat.de/images/OSCATBasic/oscat_basic333_en.pdf#page=208 *)
	VAR_INPUT
		IN : BOOL;
		PT1 : TIME;
		PTD : TIME;
		RST : BOOL;
	END_VAR
	VAR_OUTPUT
		Q : BOOL;
		W : BOOL;
	END_VAR
	VAR
		tx : TIME;
		start : TIME;
		ix : BOOL;
	END_VAR
END_FUNCTION_BLOCK

FUNCTION_BLOCK TP_X (* Generators *) (* http://www.oscat.de/images/OSCATBasic/oscat_basic333_en.pdf#page=208 *)
	VAR_INPUT
		IN : BOOL;
		PT : TIME;
	END_VAR
	VAR_OUTPUT
		Q : BOOL;
		ET : TIME;
	END_VAR
	VAR
		edge_ : BOOL;
		start : TIME;
		tx : TIME;
	END_VAR
END_FUNCTION_BLOCK

FUNCTION_BLOCK TREND (* Signal processing *) (* http://www.oscat.de/images/OSCATBasic/oscat_basic333_en.pdf#page=305 *)
	VAR_INPUT
		X : REAL;
	END_VAR
	VAR_OUTPUT
		Q : BOOL;
		TU : BOOL;
		TD : BOOL;
		D : REAL;
	END_VAR
	VAR
		last_X : REAL;
	END_VAR
END_FUNCTION_BLOCK

FUNCTION_BLOCK TREND_DW (* Signal processing *) (* http://www.oscat.de/images/OSCATBasic/oscat_basic333_en.pdf#page=315 *)
	VAR_INPUT
		X : DWORD;
	END_VAR
	VAR_OUTPUT
		Q : BOOL;
		TU : BOOL;
		TD : BOOL;
		D : DWORD;
	END_VAR
	VAR
		last_X : UDINT;
	END_VAR
END_FUNCTION_BLOCK

FUNCTION TRIANGLE_A : REAL (* Geometry *) (* http://www.oscat.de/images/OSCATBasic/oscat_basic333_en.pdf#page=107 *)
	VAR_INPUT
		S1 : REAL;
		A : REAL;
		S2 : REAL;
		S3 : REAL;
	END_VAR
END_FUNCTION

FUNCTION TRIM : BOOL (* String *) (* http://www.oscat.de/images/OSCATBasic/oscat_basic333_en.pdf#page=181 *)
	VAR_INPUT
		STR : STRING[STRING_LENGTH];
	END_VAR
	VAR_IN_OUT
		RETVAL : STRING[STRING_LENGTH]; (*Return value of the function*)
	END_VAR
	VAR
		pos : INT;
	END_VAR
END_FUNCTION

FUNCTION TRIM1 : BOOL (* String *) (* http://www.oscat.de/images/OSCATBasic/oscat_basic333_en.pdf#page=181 *)
	VAR_INPUT
		STR : STRING[STRING_LENGTH];
	END_VAR
	VAR_IN_OUT
		RETVAL : STRING[STRING_LENGTH]; (*Return value of the function*)
	END_VAR
	VAR
		pos : INT;
	END_VAR
END_FUNCTION

FUNCTION TRIME : BOOL (* String *) (* http://www.oscat.de/images/OSCATBasic/oscat_basic333_en.pdf#page=181 *)
	VAR_INPUT
		STR : STRING[STRING_LENGTH];
	END_VAR
	VAR_IN_OUT
		RETVAL : STRING[STRING_LENGTH]; (*Return value of the function*)
	END_VAR
END_FUNCTION

FUNCTION_BLOCK TUNE (* Automation *) (* http://www.oscat.de/images/OSCATBasic/oscat_basic333_en.pdf#page=472 *)
	VAR_INPUT
		SET : BOOL;
		SU : BOOL;
		SD : BOOL;
		RST : BOOL;
		SS : REAL := 0.1;
		LIMIT_L : REAL;
		LIMIT_H : REAL := 100;
		RST_VAL : REAL;
		SET_VAL : REAL := 100;
		T1 : TIME := TIME#500ms;
		T2 : TIME := TIME#2s0ms;
		S1 : REAL := 2;
		S2 : REAL := 10;
	END_VAR
	VAR_OUTPUT
		Y : REAL;
	END_VAR
	VAR
		tx : UDINT;
		start : UDINT;
		start2 : UDINT;
		state : INT;
		in : BOOL;
		step : REAL;
		SPEED : REAL;
		Y_start : REAL;
		Y_start2 : REAL;
	END_VAR
END_FUNCTION_BLOCK

FUNCTION_BLOCK TUNE2 (* Automation *) (* http://www.oscat.de/images/OSCATBasic/oscat_basic333_en.pdf#page=475 *)
	VAR_INPUT
		SET : BOOL;
		SU : BOOL;
		SD : BOOL;
		FU : BOOL;
		FD : BOOL;
		RST : BOOL;
		SS : REAL := 0.1;
		FS : REAL := 5;
		LIMIT_L : REAL;
		LIMIT_H : REAL := 100;
		RST_VAL : REAL;
		SET_VAL : REAL := 100;
		TR : TIME := TIME#500ms;
		S1 : REAL := 2;
		S2 : REAL := 10;
	END_VAR
	VAR_OUTPUT
		Y : REAL;
	END_VAR
	VAR
		tx : UDINT;
		start : UDINT;
		state : INT;
		in : BOOL;
		step : REAL;
		SPEED : REAL;
		Y_start : REAL;
	END_VAR
END_FUNCTION_BLOCK

FUNCTION T_PLC_MS : UDINT (* Measurements *) (* http://www.oscat.de/images/OSCATBasic/oscat_basic333_en.pdf#page=348 *)
	VAR CONSTANT
		debug : BOOL := 0;
		N : INT := 0;
		offset : UDINT := 0;
	END_VAR
	VAR
		tx : TIME;
	END_VAR
END_FUNCTION

FUNCTION T_PLC_US : UDINT (* Measurements *) (* http://www.oscat.de/images/OSCATBasic/oscat_basic333_en.pdf#page=351 *)
	VAR CONSTANT
		debug : BOOL := 0;
		N : INT := 0;
		offset : UDINT := 0;
	END_VAR
	VAR
		tx : TIME;
	END_VAR
END_FUNCTION

FUNCTION UPPERCASE : BOOL (* String *) (* http://www.oscat.de/images/OSCATBasic/oscat_basic333_en.pdf#page=182 *)
	VAR_INPUT
		STR : STRING[STRING_LENGTH];
	END_VAR
	VAR_IN_OUT
		RETVAL : STRING[STRING_LENGTH]; (*Return value of the function*)
	END_VAR
	VAR
		pt : REFERENCE TO BYTE;
		pos : INT;
		l : INT;
	END_VAR
END_FUNCTION

FUNCTION UTC_TO_LTIME : DATE_AND_TIME (* Time and date *) (* http://www.oscat.de/images/OSCATBasic/oscat_basic333_en.pdf#page=142 *)
	VAR_INPUT
		UTC : DATE_AND_TIME;
		DST_ENABLE : BOOL;
		TIME_ZONE_OFFSET : INT;
	END_VAR
	VAR
		tmp : INT;
	END_VAR
END_FUNCTION

FUNCTION V3_ABS : REAL (* Vector math *) (* http://www.oscat.de/images/OSCATBasic/oscat_basic333_en.pdf#page=108 *)
	VAR_INPUT
		A : VECTOR_3;
	END_VAR
END_FUNCTION

FUNCTION V3_ADD : BOOL (* Vector math *) (* http://www.oscat.de/images/OSCATBasic/oscat_basic333_en.pdf#page=108 *)
	VAR_INPUT
		A : VECTOR_3;
		B : VECTOR_3;
	END_VAR
	VAR_IN_OUT
		RETVAL : VECTOR_3; (*Return value of the function*)
	END_VAR
END_FUNCTION

FUNCTION V3_ANG : REAL (* Vector math *) (* http://www.oscat.de/images/OSCATBasic/oscat_basic333_en.pdf#page=109 *)
	VAR_INPUT
		A : VECTOR_3;
		B : VECTOR_3;
	END_VAR
	VAR
		d : REAL;
	END_VAR
END_FUNCTION

FUNCTION V3_DPRO : REAL (* Vector math *) (* http://www.oscat.de/images/OSCATBasic/oscat_basic333_en.pdf#page=109 *)
	VAR_INPUT
		A : VECTOR_3;
		B : VECTOR_3;
	END_VAR
END_FUNCTION

FUNCTION V3_NORM : BOOL (* Vector math *) (* http://www.oscat.de/images/OSCATBasic/oscat_basic333_en.pdf#page=110 *)
	VAR_INPUT
		A : VECTOR_3;
	END_VAR
	VAR_IN_OUT
		RETVAL : VECTOR_3; (*Return value of the function*)
	END_VAR
	VAR
		la : REAL;
	END_VAR
END_FUNCTION

FUNCTION V3_NUL : BOOL (* Vector math *) (* http://www.oscat.de/images/OSCATBasic/oscat_basic333_en.pdf#page=110 *)
	VAR_INPUT
		A : VECTOR_3;
	END_VAR
END_FUNCTION

FUNCTION V3_PAR : BOOL (* Vector math *) (* http://www.oscat.de/images/OSCATBasic/oscat_basic333_en.pdf#page=110 *)
	VAR_INPUT
		A : VECTOR_3;
		B : VECTOR_3;
	END_VAR
	VAR
		temp : VECTOR_3;
	END_VAR
END_FUNCTION

FUNCTION V3_REV : BOOL (* Vector math *) (* http://www.oscat.de/images/OSCATBasic/oscat_basic333_en.pdf#page=111 *)
	VAR_INPUT
		A : VECTOR_3;
	END_VAR
	VAR_IN_OUT
		RETVAL : VECTOR_3; (*Return value of the function*)
	END_VAR
END_FUNCTION

FUNCTION V3_SMUL : BOOL (* Vector math *) (* http://www.oscat.de/images/OSCATBasic/oscat_basic333_en.pdf#page=111 *)
	VAR_INPUT
		A : VECTOR_3;
		M : REAL;
	END_VAR
	VAR_IN_OUT
		RETVAL : VECTOR_3; (*Return value of the function*)
	END_VAR
END_FUNCTION

FUNCTION V3_SUB : BOOL (* Vector math *) (* http://www.oscat.de/images/OSCATBasic/oscat_basic333_en.pdf#page=112 *)
	VAR_INPUT
		A : VECTOR_3;
		B : VECTOR_3;
	END_VAR
	VAR_IN_OUT
		RETVAL : VECTOR_3; (*Return value of the function*)
	END_VAR
END_FUNCTION

FUNCTION V3_XANG : REAL (* Vector math *) (* http://www.oscat.de/images/OSCATBasic/oscat_basic333_en.pdf#page=112 *)
	VAR_INPUT
		A : VECTOR_3;
	END_VAR
	VAR
		la : REAL;
	END_VAR
END_FUNCTION

FUNCTION V3_XPRO : BOOL (* Vector math *) (* http://www.oscat.de/images/OSCATBasic/oscat_basic333_en.pdf#page=112 *)
	VAR_INPUT
		A : VECTOR_3;
		B : VECTOR_3;
	END_VAR
	VAR_IN_OUT
		RETVAL : VECTOR_3; (*Return value of the function*)
	END_VAR
END_FUNCTION

FUNCTION V3_YANG : REAL (* Vector math *) (* http://www.oscat.de/images/OSCATBasic/oscat_basic333_en.pdf#page=113 *)
	VAR_INPUT
		A : VECTOR_3;
	END_VAR
	VAR
		la : REAL;
	END_VAR
END_FUNCTION

FUNCTION V3_ZANG : REAL (* Vector math *) (* http://www.oscat.de/images/OSCATBasic/oscat_basic333_en.pdf#page=113 *)
	VAR_INPUT
		A : VECTOR_3;
	END_VAR
	VAR
		la : REAL;
	END_VAR
END_FUNCTION

FUNCTION WEEKDAY_TO_STRING : BOOL (* String *) (* http://www.oscat.de/images/OSCATBasic/oscat_basic333_en.pdf#page=182 *)
	VAR_INPUT
		WDAY : INT;
		LANG : INT;
		LX : INT;
	END_VAR
	VAR_IN_OUT
		RETVAL : STRING[10]; (*Return value of the function*)
	END_VAR
	VAR
		ly : INT;
	END_VAR
	VAR CONSTANT
		cWEEKDAYS : ARRAY[1..3,1..7] OF STRING[10] := ['Monday','Tuesday','Wednesday','Thursday','Friday','Saturday','Sunday','Montag','Dienstag','Mittwoch','Donnerstag','Freitag','Samstag','Sonntag','Lundi','Mardi','Mercredi','Jeudi','Vendredi','Samedi','Dimanche'];
		cWEEKDAYS2 : ARRAY[1..3,1..7] OF STRING[2] := ['Mo','Tu','We','Th','Fr','Sa','Su','Mo','Di','Mi','Do','Fr','Sa','So','Lu','Ma','Me','Je','Ve','Sa','Di'];
	END_VAR
END_FUNCTION

FUNCTION WINDOW : BOOL (* Mathematical *) (* http://www.oscat.de/images/OSCATBasic/oscat_basic333_en.pdf#page=69 *)
	VAR_INPUT
		LOW : REAL;
		IN : REAL;
		HIGH : REAL;
	END_VAR
END_FUNCTION

FUNCTION WINDOW2 : BOOL (* Mathematical *) (* http://www.oscat.de/images/OSCATBasic/oscat_basic333_en.pdf#page=69 *)
	VAR_INPUT
		LOW : REAL;
		IN : REAL;
		HIGH : REAL;
	END_VAR
END_FUNCTION

FUNCTION WORD_OF_BYTE : WORD (* Gate logic *) (* http://www.oscat.de/images/OSCATBasic/oscat_basic333_en.pdf#page=234 *)
	VAR_INPUT
		B1 : BYTE;
		B0 : BYTE;
	END_VAR
END_FUNCTION

FUNCTION WORD_OF_DWORD : WORD (* Gate logic *) (* http://www.oscat.de/images/OSCATBasic/oscat_basic333_en.pdf#page=235 *)
	VAR_INPUT
		IN : DWORD;
		N : BYTE;
	END_VAR
END_FUNCTION

FUNCTION WORD_TO_RANGE : REAL (* Signal processing *) (* http://www.oscat.de/images/OSCATBasic/oscat_basic333_en.pdf#page=316 *)
	VAR_INPUT
		X : WORD;
		LOW : REAL;
		HIGH : REAL;
	END_VAR
END_FUNCTION

FUNCTION WORK_WEEK : INT (* Time and date *) (* http://www.oscat.de/images/OSCATBasic/oscat_basic333_en.pdf#page=142 *)
	VAR_INPUT
		IDATE : DATE;
	END_VAR
	VAR
		d1 : DATE;
		w1 : INT;
		ds : UDINT;
		yr : INT;
		w31 : INT;
		w01 : INT;
		wm : INT;
	END_VAR
END_FUNCTION

FUNCTION YEAR_BEGIN : DATE (* Time and date *) (* http://www.oscat.de/images/OSCATBasic/oscat_basic333_en.pdf#page=143 *)
	VAR_INPUT
		Y : INT;
	END_VAR
END_FUNCTION

FUNCTION YEAR_END : DATE (* Time and date *) (* http://www.oscat.de/images/OSCATBasic/oscat_basic333_en.pdf#page=143 *)
	VAR_INPUT
		Y : INT;
	END_VAR
END_FUNCTION

FUNCTION YEAR_OF_DATE : INT (* Time and date *) (* http://www.oscat.de/images/OSCATBasic/oscat_basic333_en.pdf#page=144 *)
	VAR_INPUT
		IDATE : DATE;
	END_VAR
END_FUNCTION

FUNCTION _ARRAY_ABS : BOOL (* Array *) (* http://www.oscat.de/images/OSCATBasic/oscat_basic333_en.pdf#page=71 *)
	VAR_INPUT
		PT : REFERENCE TO ARRAY[0..32000] OF REAL;
		SIZE : UINT;
	END_VAR
	VAR
		i : UINT;
		stop : UINT;
	END_VAR
END_FUNCTION

FUNCTION _ARRAY_ADD : BOOL (* Array *) (* http://www.oscat.de/images/OSCATBasic/oscat_basic333_en.pdf#page=71 *)
	VAR_INPUT
		PT : REFERENCE TO ARRAY[0..32000] OF REAL;
		SIZE : UINT;
		X : REAL;
	END_VAR
	VAR
		i : UINT;
		stop : UINT;
	END_VAR
END_FUNCTION

FUNCTION _ARRAY_INIT : BOOL (* Array *) (* http://www.oscat.de/images/OSCATBasic/oscat_basic333_en.pdf#page=72 *)
	VAR_INPUT
		PT : REFERENCE TO ARRAY[0..32000] OF REAL;
		SIZE : UINT;
		INIT : REAL;
	END_VAR
	VAR
		i : UINT;
		stop : UINT;
	END_VAR
END_FUNCTION

FUNCTION _ARRAY_MEDIAN : REAL (* Array *) (* http://www.oscat.de/images/OSCATBasic/oscat_basic333_en.pdf#page=73 *)
	VAR_INPUT
		PT : REFERENCE TO ARRAY[0..32000] OF REAL;
		SIZE : UINT;
	END_VAR
	VAR
		i : UINT;
		stop : UINT;
	END_VAR
END_FUNCTION

FUNCTION _ARRAY_MUL : BOOL (* Array *) (* http://www.oscat.de/images/OSCATBasic/oscat_basic333_en.pdf#page=73 *)
	VAR_INPUT
		PT : REFERENCE TO ARRAY[0..32000] OF REAL;
		SIZE : UINT;
		X : REAL;
	END_VAR
	VAR
		i : UINT;
		stop : UINT;
	END_VAR
END_FUNCTION

FUNCTION _ARRAY_SHUFFLE : BOOL (* Array *) (* http://www.oscat.de/images/OSCATBasic/oscat_basic333_en.pdf#page=74 *)
	VAR_INPUT
		PT : REFERENCE TO ARRAY[0..32000] OF REAL;
		SIZE : UINT;
	END_VAR
	VAR
		temp : REAL;
		pos : INT;
		i : INT;
		stop : INT;
	END_VAR
END_FUNCTION

FUNCTION _ARRAY_SORT : BOOL (* Array *) (* http://www.oscat.de/images/OSCATBasic/oscat_basic333_en.pdf#page=75 *)
	VAR_INPUT
		PT : REFERENCE TO ARRAY[1..32000] OF REAL;
		SIZE : UINT;
	END_VAR
	VAR
		stack_count : UINT; (* Laufvariable Stack*)
		stack : ARRAY[1..32] OF UINT; (* Stackgröße~ 1,6*Log(n)/log(2) *)
		links : UINT; (* Anfangselement des Arrays *)
		rechts : UINT; (* Endelement des Arrays *)
		pivot : REAL; (* temporärer Schwellwert für Tauschbedingung *)
		i : UINT; (* Laufvariable1 *)
		j : UINT; (* Laufvariable2 *)
		ende_innen : BOOL; (* Ende innere Schleife *)
		ende_aussen : BOOL; (* Ende äußere Schleife *)
		tmp : REAL; (* Hilfsvariable zum Tauschen von Werten *)
	END_VAR
END_FUNCTION

FUNCTION _BUFFER_CLEAR : BOOL (* Buffer Management *) (* http://www.oscat.de/images/OSCATBasic/oscat_basic333_en.pdf#page=477 *)
	VAR_INPUT
		PT : REFERENCE TO BYTE;
		SIZE : UINT;
	END_VAR
	VAR
		ptw : REFERENCE TO DWORD;
		temp : UDINT;
		end : UDINT;
		end32 : UDINT;
	END_VAR
END_FUNCTION

FUNCTION _BUFFER_INIT : BOOL (* Buffer Management *) (* http://www.oscat.de/images/OSCATBasic/oscat_basic333_en.pdf#page=477 *)
	VAR_INPUT
		PT : REFERENCE TO BYTE;
		SIZE : UINT;
		INIT : BYTE;
	END_VAR
	VAR
		ptw : REFERENCE TO DWORD;
		temp : UDINT;
		end : UDINT;
		end32 : UDINT;
	END_VAR
END_FUNCTION

FUNCTION _BUFFER_INSERT : INT (* Buffer Management *) (* http://www.oscat.de/images/OSCATBasic/oscat_basic333_en.pdf#page=478 *)
	VAR_INPUT
		STR : STRING[STRING_LENGTH];
		POS : INT;
		PT : REFERENCE TO ARRAY[0..32767] OF BYTE;
		SIZE : UINT;
	END_VAR
	VAR
		end : INT;
		lx : INT;
		i : INT;
	END_VAR
END_FUNCTION

FUNCTION _BUFFER_UPPERCASE : BOOL (* Buffer Management *) (* http://www.oscat.de/images/OSCATBasic/oscat_basic333_en.pdf#page=479 *)
	VAR_INPUT
		PT : REFERENCE TO ARRAY[0..32000] OF BYTE;
		SIZE : INT;
	END_VAR
	VAR
		pos : INT;
	END_VAR
END_FUNCTION

FUNCTION_BLOCK _RMP_B (* Signal generators *) (* http://www.oscat.de/images/OSCATBasic/oscat_basic333_en.pdf#page=255 *)
	VAR_INPUT
		DIR : BOOL; (* true = up *)
		E : BOOL := TRUE;
		TR : TIME;
	END_VAR
	VAR_IN_OUT
		RMP : BYTE;
	END_VAR
	VAR
		tx : TIME;
		tl : TIME;
		tn : TIME;
		init : BOOL;
		last_dir : BOOL;
		start : BYTE;
	END_VAR
END_FUNCTION_BLOCK

FUNCTION_BLOCK _RMP_NEXT (* Signal generators *) (* http://www.oscat.de/images/OSCATBasic/oscat_basic333_en.pdf#page=255 *)
	VAR_INPUT
		E : BOOL := TRUE;
		IN : BYTE;
		TR : TIME;
		TF : TIME;
		TL : TIME;
	END_VAR
	VAR_OUTPUT
		DIR : BOOL; (* upwards = TRUE *)
		UP : BOOL;
		DN : BOOL;
	END_VAR
	VAR_IN_OUT
		OUT : BYTE;
	END_VAR
	VAR
		rmx : _RMP_B;
		dirx : TREND_DW;
		t_lock : TP;
		xen : BOOL;
		xdir : BOOL;
	END_VAR
END_FUNCTION_BLOCK

FUNCTION_BLOCK _RMP_W (* Signal generators *) (* http://www.oscat.de/images/OSCATBasic/oscat_basic333_en.pdf#page=256 *)
	VAR_INPUT
		DIR : BOOL;
		E : BOOL := TRUE;
		TR : TIME;
	END_VAR
	VAR_IN_OUT
		RMP : WORD;
	END_VAR
	VAR
		tx : UDINT;
		tl : UDINT;
		step : DINT;
		init : BOOL;
		last_dir : BOOL;
	END_VAR
END_FUNCTION_BLOCK

FUNCTION _STRING_TO_BUFFER : INT (* Buffer Management *) (* http://www.oscat.de/images/OSCATBasic/oscat_basic333_en.pdf#page=479 *)
	VAR_INPUT
		STR : STRING[STRING_LENGTH];
		POS : INT;
		PT : REFERENCE TO ARRAY[0..32767] OF BYTE;
		SIZE : UINT;
	END_VAR
	VAR
		ps : REFERENCE TO BYTE;
		i : INT;
		end : INT;
	END_VAR
END_FUNCTION

(* ---- PARSET.st ---- *)
FUNCTION_BLOCK PARSET
    (*http://www.oscat.de/images/OSCATBasic/oscat_basic333_en.pdf#page=466*)
    (* read system_time *)
    tx := T_PLC_MS();

    (* init sequence *)
    IF NOT init THEN
    	set.0 := NOT A0;
    	init := TRUE;
    	X[0,1] := X01;
    	X[0,2] := X02;
    	X[0,3] := X03;
    	X[0,4] := X04;
    	X[1,1] := X11;
    	X[1,2] := X12;
    	X[1,3] := X13;
    	X[1,4] := X14;
    	X[2,1] := X21;
    	X[2,2] := X22;
    	X[2,3] := X23;
    	X[2,4] := X24;
    	X[3,1] := X31;
    	X[3,2] := X32;
    	X[3,3] := X33;
    	X[3,4] := X34;
    	P1 := X01;
    	P2 := X02;
    	P3 := X03;
    	P4 := X04;
    END_IF

    (* check for input change *)
    IF (A0 XOR set.0) OR (A1 XOR set.1) THEN
    	(* a new set is selected *)
    	set.0 := A0;
    	set.1 := A1;
    	IF TC > t#0s THEN
    		start := TRUE;
    		last := tx;
    		(* save the step speed for the output changes in S *)
    		S1 := (X[set,1] - P1)/UDINT_TO_REAL(TIME_TO_UDINT(TC));
    		S2 := (X[set,2] - P2)/UDINT_TO_REAL(TIME_TO_UDINT(TC));
    		S3 := (X[set,3] - P3)/UDINT_TO_REAL(TIME_TO_UDINT(TC));
    		S4 := (X[set,4] - P4)/UDINT_TO_REAL(TIME_TO_UDINT(TC));
    	END_IF
    ELSIF start AND tx - last < TIME_TO_UDINT(TC) THEN
    	(* ramp the outputs to the new value *)
    	P1 := X[set,1] - S1 * UDINT_TO_REAL(TIME_TO_UDINT(TC) - tx + last);
    	P2 := X[set,2] - S2 * UDINT_TO_REAL(TIME_TO_UDINT(TC) - tx + last);
    	P3 := X[set,3] - S3 * UDINT_TO_REAL(TIME_TO_UDINT(TC) - tx + last);
    	P4 := X[set,4] - S4 * UDINT_TO_REAL(TIME_TO_UDINT(TC) - tx + last);
    ELSE
    	(* make sure outputs match the correct set values *)
    	start := FALSE;
    	P1 := X[set,1];
    	P2 := X[set,2];
    	P3 := X[set,3];
    	P4 := X[set,4];
    END_IF

    (* revision history
    hm	2.11.2007		rev 1.0
    	original version

    hm	16. mar. 2008	rev 1.1
    	added type conversions to avoid warnings under codesys 3.0

    *)

END_FUNCTION_BLOCK

(* ---- PARSET2.st ---- *)
FUNCTION_BLOCK PARSET2
    (*http://www.oscat.de/images/OSCATBasic/oscat_basic333_en.pdf#page=467*)
    (* init sequence *)
    IF NOT init THEN
    	init := TRUE;
    	Pset(TC:=TC, X01:=X01, X02:=X02, X03:=X03, X04:=X04, X11:=X11, X12:=X12, X13:=X13, X14:=X14, X21:=X21, X22:=X22, X23:=X23, X24:=X24, X31:=X31, X32:=X32, X33:=X33, X34:=X34);
    END_IF
    IF ABS(X) < L1 THEN
    	Pset(A0 := FALSE, A1 := FALSE);
    ELSIF ABS(X) < L2 THEN
    	Pset(A0 := TRUE, A1 := FALSE);
    ELSIF ABS(X) < L3 THEN
    	Pset(A0 := FALSE, A1 := TRUE);
    ELSE
    	Pset(A0 := TRUE, A1 := TRUE);
    END_IF
    P1 := Pset.P1;
    P2 := Pset.P2;
    P3 := Pset.P3;
    P4 := Pset.P4;

    (* revision history
    hm		3.11.2007		rev 1.0
    	original version

    *)

END_FUNCTION_BLOCK

(* ---- PIN_CODE.st ---- *)
FUNCTION_BLOCK PIN_CODE
    (*http://www.oscat.de/images/OSCATBasic/oscat_basic333_en.pdf#page=231*)
    TP := FALSE;
    IF E THEN
    	IF CB = CODE(PIN, POS) THEN
    		POS := POS + 1;
    		IF POS > LEN(PIN) THEN
    			(* proper code is detected *)
    			TP := TRUE;
    			POS := 1;
    		END_IF
    	ELSE
    		POS := 1;
    	END_IF
    END_IF

    (* revision history
    hm	30. oct. 2008	rev 1.0
    	original version

    *)

END_FUNCTION_BLOCK

(* ---- PRESSURE.st ---- *)
FUNCTION_BLOCK PRESSURE
    (*http://www.oscat.de/images/OSCATBasic/oscat_basic333_en.pdf#page=371*)
    YBAR := BAR +
    		PA * 1.0E-5 +
    		0.980665 * ATT +
    		1.01325 * ATM +
    		0.001333224 * TORR +
    		0.0980665 * MWS;
    YMWS := YBAR * 10.1971621297793;
    YTORR := YBAR * 750.0615050434140;
    YATT := YBAR * 1.0197162129779;
    YATM := YBAR * 0.9869232667160;
    YPA := YBAR * 100000.0;

    (*
    Druck, Pascal PA 1 PA = 1 N/m2 = 1 kg/(s2 E m) . 0,75 E 10.2 mmHg
    mechanische 1 MPa = 1 N/mm2 . fur Festigkeitsangaben
    Spannung BAR BAR 1 BAR = 105 PA = 103 mbar = 105 kg/(s2 E m)
    Millimeter- mmHg 1 mmHg = 133,322 PA = 1,333 22 mbar
    Quecksilbersaule . nur in Heilkunde zulassig
    physik. Atmosphare ATM 1 ATM = 1,013 25 BAR
    techn. Atmosphare at 1 at = 1 kp/cm2 = 0,980665 BAR
    TORR TORR 1 TORR = (101325/760) PA = 1,333224 mbar
    Meter-Wassersaule MWS 1 MWS = 9806,65 PA = 98,0665 mbar
    psi lbf/in2 1 lbf/in2 = 68,947 57 mbar = 6894,757 PA

    *)

    (* revision history

    hm	27. mar. 2007	rev 1.0
    	original version

    hm	11. mar. 2009	rev 1.1
    	improved code

    *)
END_FUNCTION_BLOCK

(* ---- PWM_DC.st ---- *)
FUNCTION_BLOCK PWM_DC
    (*http://www.oscat.de/images/OSCATBasic/oscat_basic333_en.pdf#page=263*)
    IF F > 0.0 THEN
    	tmp := 1000.0 / F;
    	clk(PT := REAL_TO_TIME(tmp));
    	pulse(IN := clk.Q, PT := REAL_TO_TIME(tmp * DC));
    	Q := pulse.Q;
    END_IF

    (* revision history

    hm	25. feb 2007	rev 1.1
    	recoded in st for better performance and better portability

    hm	27. nov 2007	rev 1.2
    	avoid divide by 0 when F = 0

    hm	19. oct. 2008	rev 1.3
    	changed type TP_R to TP_X because of name change
    	improved performance

    hm	11. mar. 2009	rev 1.4
    	changed real constants to use dot syntax

    *)
END_FUNCTION_BLOCK

(* ---- PWM_PW.st ---- *)
FUNCTION_BLOCK PWM_PW
    (*http://www.oscat.de/images/OSCATBasic/oscat_basic333_en.pdf#page=264*)
    IF F > 0.0 THEN
    	clk(PT := REAL_TO_TIME(1000.0 / F));
    	pulse(IN := clk.Q, PT := PW);
    	Q := pulse.Q;
    END_IF

    (* revision history

    hm	25. feb 2007	rev 1.1
    	recoded in st for better performance and better portability

    hm	27. nov 2007	rev 1.2
    	avoid divide by 0 when F = 0

    hm	9. dec 2007		rev 1.3
    	corrected an error with F = 0

    hm	19. oct. 2008	rev 1.4
    	changed type tp_r to TP_x brecause of name change

    hm	11. mar. 2009	rev 1.5
    	changed real constants to use dot syntax

    *)
END_FUNCTION_BLOCK

(* ---- RMP_B.st ---- *)
FUNCTION_BLOCK RMP_B
    (*http://www.oscat.de/images/OSCATBasic/oscat_basic333_en.pdf#page=264*)
    (* generate ramp *)
    rmp(DIR := UP, E := E, TR := PT, RMP := OUT);

    (* SET or reset operation *)
    IF RST THEN
    	OUT := 0;
    ELSIF SET THEN
    	OUT := 255;
    END_IF

    (* checks for outputs stable and reset or SET BUSY flag *)
    LOW := OUT = 0;
    HIGH := OUT = 255;
    BUSY := NOT (LOW OR HIGH) AND E;

    (* revision history

    hm 5.10.2006	rev 1.1
    	added BUSY output
    hm 17.1.2007	rev 1.2
    	renamed input ud to UP for better usability
    	deleted unused variable step

    hm	17.9.2007		rev 1.3
    	replaced time() with t_plc_ms() for compatibility reasons

    hm	28. sep 2007	rev 1.4
    	added outputs on and off
    	BUSY is now disabled while en is false
    	new coding for higher accuracy and performance

    hm	5. oct 2007	rev 1.5
    	added statements to allow for PT to be t#0s output jumps to max or min immediately

    hm	25. dec 2007	rev 1.6
    	improved code for better performance

    hm	16. oct. 2008	rev 1.7
    	improved code for better performance

    hm	18. oct. 2008	rev 1.8
    	added type conversion to avoid warnings
    	changed input en to E for compatibility reasons

    hm	23. oct. 2008	REV 	2.0
    	new code using _RMP_B

    *)
END_FUNCTION_BLOCK

(* ---- RMP_SOFT.st ---- *)
FUNCTION_BLOCK RMP_SOFT
    (*http://www.oscat.de/images/OSCATBasic/oscat_basic333_en.pdf#page=266*)
    tmp := SEL(IN, 0, VAL);
    IF tmp > OUT THEN
    	(* we need to ramp down *)
    	rmp(DIR := TRUE, E := TRUE, TR := PT_ON, RMP := OUT);
    	(* make sure OUT does not surpass tmp *)
    	OUT := MIN(OUT, tmp);
    ELSIF tmp < OUT THEN
    	(* we need to ramp up *)
    	rmp(DIR := FALSE, E := TRUE, TR := PT_OFF, RMP := OUT);
    	(* make sure OUT does not surpass tmp *)
    	OUT := MAX(OUT, tmp);
    ELSE
    	(* no ramp necessary *)
    	rmp(E := FALSE, RMP := OUT);
    END_IF

    (* revision history

    hm 22.1.2007	rev 1.1
    	deleted unused variables X1 and I, X2 and X3

    hm	17.9.2007	rev 1.2
    	replaced time() with t_plc_ms() for compatibility reasons

    hm	26. oct. 2008	2.0
    	new code using _rmp_b
    *)

END_FUNCTION_BLOCK

(* ---- RMP_W.st ---- *)
FUNCTION_BLOCK RMP_W
    (*http://www.oscat.de/images/OSCATBasic/oscat_basic333_en.pdf#page=267*)
    (* generate ramp *)
    rmp(DIR := UP, E := E, TR := PT, RMP := OUT);

    (* SET or reset operation *)
    IF RST THEN
    	OUT := 0;
    ELSIF SET THEN
    	OUT := 65535;
    END_IF

    (* checks for outputs stable and reset or SET BUSY flag *)
    LOW := OUT = 0;
    HIGH := OUT = 65535;
    BUSY := NOT (LOW OR HIGH) AND E;

    (* revision history:

    hm 4.10.2006		rev 1.1
    	added the BUSY output which signals that the ramp is running.

    hm 22.1.2007		rev 1.2
    	deleted unused variable step

    hm	17.9.2007		rev 1.3
    	replaced time() with t_plc_ms() for compatibility reasons

    hm	28. sep 2007	rev 1.4
    	added outputs on and off
    	BUSY is now disabled while en is false
    	new coding for higher accuracy and performance

    hm	5. oct 2007	rev 1.5
    	added statements to allow for PT to be t#0s output jumps to max or min immediately

    hm	2. dec 2007	rev 1.6
    	corrected an error in calculation of step response

    hm	25. dec 2007	rev 1.7
    	corrected an error while step response was too slow for fast rise times

    hm	16. oct. 2008	rev 1.8
    	improved performance

    hm	18. oct. 2008	rev 1.9
    	renamed inout EN to E for compatibility reasons

    hm	23. oct. 2008	rev 2.0
    	new code using _RMP_W
    *)

END_FUNCTION_BLOCK

(* ---- RTC_2.st ---- *)
FUNCTION_BLOCK RTC_2
    (*http://www.oscat.de/images/OSCATBasic/oscat_basic333_en.pdf#page=133*)
    (* call rtc *)
    RT(SET := SET, SDT := SDT, SMS := SMS);
    UDT := RT.XDT;
    XMS := RT.XMS;

    (* check for daylight savings time and SET DSO output *)
    DSO := DST(UDT) AND DEN;

    (* calculate time offset and SET ldt output *)
    LOCAL_DT := UDINT_TO_DT(DT_TO_UDINT(UDT) + INT_TO_UDINT(OFS + BOOL_TO_INT(DSO)*60) * 60);

    (* revision history
    hm		20. jan. 2008	rev 1.0
    	original version

    hm		20. feb. 2008	rev 1.1
    	added Millisecond SET input

    hm		12. jun. 2008	rev 1.2
    	improved performance

    hm		20. jan. 2011	rev 1.3
    	changed offset to be in minutes

    hm		27. apr. 2011	rev 1.4
    	fixed error with local time calculation

    hm     3. Feb 2021     rev 1.5
         changed LDT to LOCAL_DT for compatibility with IEC61131-3

    *)
END_FUNCTION_BLOCK

(* ---- RTC_MS.st ---- *)
FUNCTION_BLOCK RTC_MS
    (*http://www.oscat.de/images/OSCATBasic/oscat_basic333_en.pdf#page=134*)
    Tx := T_PLC_MS();
    IF SET OR NOT init THEN
    	(* clock needs to be SET when SET is true or after power up *)
    	init := TRUE;
    	XDT := SDT;
    	XMS := SMS;
    ELSE
    	XMS := XMS + UDINT_TO_INT(Tx - last);
    	(* check if one second has expired *)
    	IF XMS > 999 THEN
    		XDT := XDT + T#1s;
    		XMS := XMS - 1000;
    	END_IF
    END_IF
    last := Tx;

    (* revision history
    hm		20. jan. 2008	rev 1.0
    	original version

    hm		20. feb. 2008	rev 1.1
    	added Millisecond SET input
    *)
END_FUNCTION_BLOCK

(* ---- SCHEDULER.st ---- *)
FUNCTION_BLOCK SCHEDULER
    (*http://www.oscat.de/images/OSCATBasic/oscat_basic333_en.pdf#page=198*)
    (* read system_time *)
    tx := UDINT_TO_TIME(T_PLC_MS());

    IF NOT init THEN
    	init := TRUE;
    	s0 := tx - T0;
    	s1 := tx - T1;
    	s2 := tx - T2;
    	s3 := tx - T3;
    END_IF

    Q0 := FALSE;
    Q1 := FALSE;
    Q2 := FALSE;
    Q3 :=FALSE;

    CASE c OF
    	0: 	IF tx - s0 >= T0 THEN
    			Q0 := E0;
    			s0 := tx;
    		END_IF
    		c := 1;
    	1: 	IF tx - s1 >= T1 THEN
    			Q1 := E1;
    			s1 := tx;
    		END_IF
    		c := 2;
    	2: 	IF tx - s2 >= T2 THEN
    			Q2 := E2;
    			s2 := tx;
    		END_IF
    		c := 3;
    	3: 	IF tx - s3 >= T3 THEN
    			Q3 := E3;
    			s3 := tx;
    		END_IF
    		c := 0;
    END_CASE

    (* revision history

    hm 28. sep. 2008	rev 1.0
    	original version

    hm	14. mar. 2009	rev 1.1
    	removed double assignments

    *)
END_FUNCTION_BLOCK

(* ---- SCHEDULER_2.st ---- *)
FUNCTION_BLOCK SCHEDULER_2
    (*http://www.oscat.de/images/OSCATBasic/oscat_basic333_en.pdf#page=198*)
    Q0 := E0 AND (sx MOD C0 - O0 = 0);
    Q1 := E1 AND (sx MOD C1 - O1 = 0);
    Q2 := E2 AND (sx MOD C2 - O2 = 0);
    Q3 := E3 AND (sx MOD C3 - O3 = 0);

    (* increment cycle counter every cycle *)
    sx := sx + 1;

    (* revision history
    hm 29. sep. 2008		rev 1.0
    	original version

    *)
END_FUNCTION_BLOCK

(* ---- SEL2_OF_3.st ---- *)
FUNCTION_BLOCK SEL2_OF_3
    (*http://www.oscat.de/images/OSCATBasic/oscat_basic333_en.pdf#page=298*)
    D12 := ABS(IN1-IN2) <= D;
    D23 := ABS(IN2-IN3) <= D;
    D31 := ABS(IN3-IN1) <= D;

    IF (D12 AND D23) OR (D12 AND D31) OR (D23 AND D31) THEN
    	(* all 3 inputs are valid *)
    	Y := (IN1 + IN2 + IN3) * 0.333333333333;
    	E := FALSE;
    	W := 0;
    ELSIF D12 THEN
    	(* only inut 1 and 2 are valid *)
    	Y := (IN1 + IN2) * 0.5;
    	E := FALSE;
    	W := 3;
    ELSIF D23 THEN
    	(* only inut 2 and 3 are valid *)
    	Y := (IN2 + IN3) * 0.5;
    	E := FALSE;
    	W := 1;
    ELSIF D31 THEN
    	(* only inut 3 and 1 are valid *)
    	Y := (IN3 + IN1) * 0.5;
    	E := FALSE;
    	W := 2;
    ELSE
    	(* no calculation possible *)
    	E := TRUE;
    	W := 4;
    END_IF

    (* revision history
    hm	18. may 2008	rev 1.0
    	original version

    hm	10. mar. 2009	rev 1.1
    	improved code
    *)
END_FUNCTION_BLOCK

(* ---- SEL2_OF_3B.st ---- *)
FUNCTION_BLOCK SEL2_OF_3B
    (*http://www.oscat.de/images/OSCATBasic/oscat_basic333_en.pdf#page=299*)
    Q := (IN1 AND IN2) OR (IN1 AND IN3) OR (IN2 AND IN3);
    TDEL(IN := (IN1 XOR IN2) OR (IN1 XOR IN3) OR (IN2 XOR IN3), PT := TD);
    W := TDEL.Q;

    (* revision history
    hm		19. may 2008	rev 1.0
    	original version

    *)
END_FUNCTION_BLOCK

(* ---- SELECT_8.st ---- *)
FUNCTION_BLOCK SELECT_8
    (*http://www.oscat.de/images/OSCATBasic/oscat_basic333_en.pdf#page=247*)
    IF RST THEN
    	STATE := 0;
    ELSIF SET THEN
    	STATE := BYTE_TO_INT(IN);
    ELSIF UP AND NOT last_up THEN
    	STATE := INC(STATE,1,7);
    ELSIF DN AND NOT last_dn THEN
    	STATE := INC(STATE,-1,7);
    END_IF
    last_up := UP;
    last_dn := DN;

    Q0 := FALSE;
    Q1 := FALSE;
    Q2 := FALSE;
    Q3 := FALSE;
    Q4 := FALSE;
    Q5 := FALSE;
    Q6 := FALSE;
    Q7 := FALSE;

    IF E THEN
    	CASE STATE OF
    		0: Q0 := TRUE;
    		1: Q1 := TRUE;
    		2: Q2 := TRUE;
    		3: Q3 := TRUE;
    		4: Q4 := TRUE;
    		5: Q5 := TRUE;
    		6: Q6 := TRUE;
    		7: Q7 := TRUE;
    	END_CASE
    END_IF

    (* revision history
    hm	16. jan 2008	rev 1.0
    	original version

    hm	27. feb. 2009	rev 1.1
    	renamed input en to E
    *)
END_FUNCTION_BLOCK

(* ---- SEQUENCE_4.st ---- *)
FUNCTION_BLOCK SEQUENCE_4
    (*http://www.oscat.de/images/OSCATBasic/oscat_basic333_en.pdf#page=199*)
    (* read sps timer *)
    tx := UDINT_TO_TIME(T_PLC_MS());

    (* initialize on startup *)
    IF NOT init THEN
    	last := tx;
    	init := TRUE;
    	STATUS := 110;
    END_IF

    (* asynchronous reset *)
    IF RST THEN
    	STEP := -1;
    	Q0 := 0;
    	Q1 := 0;
    	Q2 := 0;
    	Q3 := 0;
    	STATUS := 110;
    	RUN := 0;

    (* edge_ on START input restarts the sequencer *)
    ELSIF START AND NOT edge_ THEN
    	STEP := 0;
    	last := tx;
    	STATUS := 111;
    	Q0 := 0;
    	Q1 := 0;
    	Q2 := 0;
    	Q3 := 0;
    	RUN := 1;
    END_IF
    edge_ := START;

    (* check if stop on STATUS is necessary *)
    IF STATUS > 0 AND STATUS < 100 AND STOP_ON_ERROR THEN RETURN; END_IF

    (* sequence is running *)
    IF RUN AND STEP = 0 THEN
    	IF NOT Q0 AND IN0 AND tx - last <= WAIT0 THEN
    		Q0 := TRUE;
    		last := tx;
    	ELSIF NOT Q0 AND tx - last > WAIT0 THEN
    		STATUS := 1;
    		RUN := FALSE;
    	ELSIF Q0 AND tx - last >= DELAY0 THEN
    		STEP := 1;
    		last := tx;
    	END_IF
    END_IF
    IF RUN AND STEP = 1 THEN
    	IF NOT Q1 AND IN1 AND tx - last <= WAIT1 THEN
    		Q0 := FALSE;
    		Q1 := TRUE;
    		last := tx;
    	ELSIF NOT Q1 AND tx - last > WAIT1 THEN
    		STATUS := 2;
    		Q0 := FALSE;
    		RUN := FALSE;
    	ELSIF Q1 AND tx - last >= DELAY1 THEN
    		STEP := 2;
    		last := tx;
    	END_IF
    END_IF
    IF RUN AND STEP = 2 THEN
    	IF NOT Q2 AND IN2 AND tx - last <= WAIT2 THEN
    		Q1 := FALSE;
    		Q2 := TRUE;
    		last := tx;
    	ELSIF NOT Q2 AND tx - last > WAIT2 THEN
    		STATUS := 3;
    		Q1 := FALSE;
    		RUN := FALSE;
    	ELSIF Q2 AND tx - last >= DELAY2 THEN
    		STEP := 3;
    		last := tx;
    	END_IF
    END_IF
    IF RUN AND STEP = 3 THEN
    	IF NOT Q3 AND IN3 AND tx - last <= WAIT3 THEN
    		Q2 := FALSE;
    		Q3 := TRUE;
    		last := tx;
    	ELSIF NOT Q3 AND tx - last > WAIT3 THEN
    		STATUS := 4;
    		Q2 := FALSE;
    		RUN := FALSE;
    	ELSIF Q3 AND tx - last >= DELAY3 THEN
    		STEP := -1;
    		Q3 := FALSE;
    		RUN := FALSE;
    		STATUS := 110;
    	END_IF
    END_IF
    QX := Q0 OR Q1 OR Q2 OR Q3;

    (*
    hm 1.10.06		rev 1.1
    	corrected delay logic to be after event and not before
    	added any output

    hm 1.12.06		rev 1.2
    	corrected failure in sequence logic.
    	added init at startup to prevent from initial error after START.

    hm 17.1.2007		rev 1.3
    	changed output fault to STATUS for better compatibility with other modules (ESR).
    	added stop on error functionality and setup variable
    	default for inputs IN0..3 is true.
    	renamed variable state to STEP

    hm	17.sep 2007	rev 1.4
    	replaced time() with T_PLC_MS() for compatibility reasons

    hm	13. mar. 2009	rev 1.5
    	renamed output any to QX for compatibility resons

    *)
END_FUNCTION_BLOCK

(* ---- SEQUENCE_64.st ---- *)
FUNCTION_BLOCK SEQUENCE_64
    (*http://www.oscat.de/images/OSCATBasic/oscat_basic333_en.pdf#page=202*)
    (* read system timer *)
    tx := UDINT_TO_TIME(T_PLC_MS());
    TRIG := FALSE;

    IF RST THEN
    	STATE := -1;

    (* START sequence *)
    ELSIF START AND NOT edge_ THEN
    	STATE := 0;
    	last := tx;
    	TRIG := TRUE;

    (* sequence generator *)
    ELSIF (STATE >= 0) THEN
    	IF (tx - last) >= PROG[STATE] THEN
    		STATE := INC2(STATE, 1, -1, SMAX);
    		last := tx;
    		TRIG := TRUE;
    	END_IF
    END_IF

    edge_ := START;

    (* revision history
    hm	29. jun. 2008
    	original version

    *)
END_FUNCTION_BLOCK

(* ---- SEQUENCE_8.st ---- *)
FUNCTION_BLOCK SEQUENCE_8
    (*http://www.oscat.de/images/OSCATBasic/oscat_basic333_en.pdf#page=203*)
    (* read sps timer *)
    tx := UDINT_TO_TIME(T_PLC_MS());

    (* initialize on startup *)
    IF NOT init THEN
    	last := tx;
    	init := TRUE;
    	STATUS := 110;
    END_IF

    (* asynchronous reset *)
    IF RST THEN
    	STEP := -1;
    	Q0 := 0;
    	Q1 := 0;
    	Q2 := 0;
    	Q3 := 0;
    	Q4 := 0;
    	Q5 := 0;
    	Q6 := 0;
    	Q7 := 0;
    	STATUS := 110;
    	RUN := 0;

    (* edge_ on START input restarts the sequencer *)
    ELSIF START AND NOT edge_ THEN
    	STEP := 0;
    	last := tx;
    	STATUS := 111;
    	Q0 := 0;
    	Q1 := 0;
    	Q2 := 0;
    	Q3 := 0;
    	Q4 := 0;
    	Q5 := 0;
    	Q6 := 0;
    	Q7 := 0;
    	RUN := 1;
    END_IF
    edge_ := START;

    (* check if stop on error is necessary *)
    IF STATUS > 0 AND STATUS < 100 AND STOP_ON_ERROR THEN RETURN; END_IF

    (* sequence is running *)
    IF RUN AND STEP = 0 THEN
    	IF NOT Q0 AND IN0 AND tx - last <= WAIT0 THEN
    		Q0 := TRUE;
    		last := tx;
    	ELSIF NOT Q0 AND tx - last > WAIT0 THEN
    		STATUS := 1;
    		RUN := FALSE;
    	ELSIF Q0 AND tx - last >= DELAY0 THEN
    		STEP := 1;
    		last := tx;
    	END_IF
    END_IF
    IF RUN AND STEP = 1 THEN
    	IF NOT Q1 AND IN1 AND tx - last <= WAIT1 THEN
    		Q0 := FALSE;
    		Q1 := TRUE;
    		last := tx;
    	ELSIF NOT Q1 AND tx - last > WAIT1 THEN
    		STATUS := 2;
    		Q0 := FALSE;
    		RUN := FALSE;
    	ELSIF Q1 AND tx - last >= DELAY1 THEN
    		STEP := 2;
    		last := tx;
    	END_IF
    END_IF
    IF RUN AND STEP = 2 THEN
    	IF NOT Q2 AND IN2 AND tx - last <= WAIT2 THEN
    		Q1 := FALSE;
    		Q2 := TRUE;
    		last := tx;
    	ELSIF NOT Q2 AND tx - last > WAIT2 THEN
    		STATUS := 3;
    		Q1 := FALSE;
    		RUN := FALSE;
    	ELSIF Q2 AND tx - last >= DELAY2 THEN
    		STEP := 3;
    		last := tx;
    	END_IF
    END_IF
    IF RUN AND STEP = 3 THEN
    	IF NOT Q3 AND IN3 AND tx - last <= WAIT3 THEN
    		Q2 := FALSE;
    		Q3 := TRUE;
    		last := tx;
    	ELSIF NOT Q3 AND tx - last > WAIT3 THEN
    		STATUS := 4;
    		Q2 := FALSE;
    		RUN := FALSE;
    	ELSIF Q3 AND tx - last >= DELAY3 THEN
    		STEP := 4;
    		last := tx;
    	END_IF
    END_IF
    IF RUN AND STEP = 4 THEN
    	IF NOT Q4 AND IN4 AND tx - last <= WAIT4 THEN
    		Q3 := FALSE;
    		Q4 := TRUE;
    		last := tx;
    	ELSIF NOT Q4 AND tx - last > WAIT4 THEN
    		STATUS := 5;
    		Q3 := FALSE;
    		RUN := FALSE;
    	ELSIF Q4 AND tx - last >= DELAY4 THEN
    		STEP := 5;
    		last := tx;
    	END_IF
    END_IF
    IF RUN AND STEP = 5 THEN
    	IF NOT Q5 AND IN5 AND tx - last <= WAIT5 THEN
    		Q4 := FALSE;
    		Q5 := TRUE;
    		last := tx;
    	ELSIF NOT Q5 AND tx - last > WAIT5 THEN
    		STATUS := 6;
    		Q4 := FALSE;
    		RUN := FALSE;
    	ELSIF Q5 AND tx - last >= DELAY5 THEN
    		STEP := 6;
    		last := tx;
    	END_IF
    END_IF
    IF RUN AND STEP = 6 THEN
    	IF NOT Q6 AND IN6 AND tx - last <= WAIT6 THEN
    		Q5 := FALSE;
    		Q6 := TRUE;
    		last := tx;
    	ELSIF NOT Q6 AND tx - last > WAIT6 THEN
    		STATUS := 7;
    		Q5 := FALSE;
    		RUN := FALSE;
    	ELSIF Q6 AND tx - last >= DELAY6 THEN
    		STEP := 7;
    		last := tx;
    	END_IF
    END_IF
    IF RUN AND STEP = 7 THEN
    	IF NOT Q7 AND IN7 AND tx - last <= WAIT7 THEN
    		Q6 := FALSE;
    		Q7 := TRUE;
    		last := tx;
    	ELSIF NOT Q7 AND tx - last > WAIT7 THEN
    		STATUS := 8;
    		Q6 := FALSE;
    		RUN := FALSE;
    	ELSIF Q7 AND tx - last >= DELAY7 THEN
    		STEP := -1;
    		Q7 := FALSE;
    		RUN := FALSE;
    		STATUS := 110;
    	END_IF
    END_IF
    QX := Q0 OR Q1 OR Q2 OR Q3 OR Q4 OR Q5 OR Q6 OR Q7;

    (*
    hm 1.10.06		rev 1.1
    	corrected delay logic to be after event and not before
    	added any output

    hm 1.12.06		rev 1.2
    	corrected failure in sequence logic.
    	added init at startup to prevent from initial statuss after START.

    hm 17.1.2007		rev 1.3
    	changed output fault to STATUS for better compatibility with other modules (ESR)
    	added stop on error functionality and setup variable
    	default for inputs IN0..7 is true.
    	renames variable state to STEP

    hm	17.sep 2007	rev 1.4
    	replaced time() with T_PLC_MS() for compatibility reasons

    hm	13. mar. 2009	rev 1.5
    	renamed output any to QX for compatibility resons

    *)
END_FUNCTION_BLOCK

(* ---- SH.st ---- *)
FUNCTION_BLOCK SH
    (*http://www.oscat.de/images/OSCATBasic/oscat_basic333_en.pdf#page=299*)
    IF CLK AND NOT edge_ THEN
    	OUT := IN;
    	TRIG := TRUE;
    ELSE;
    	TRIG := FALSE;
    END_IF
    edge_ := CLK;

    (* revision history

    hm 16.1.2007	rev 1.1
    	added TRIG output

    *)
END_FUNCTION_BLOCK

(* ---- SH_1.st ---- *)
FUNCTION_BLOCK SH_1
    (*http://www.oscat.de/images/OSCATBasic/oscat_basic333_en.pdf#page=300*)
    (* read system time *)
    tx := UDINT_TO_TIME(T_PLC_MS());

    IF tx - last >= PT THEN
    	last := tx;
    	OUT := IN;
    	TRIG := TRUE;
    ELSE
    	TRIG := FALSE;
    END_IF

    (* revision history

    HM	6.1.2007	rev 1.1
    	added TRIG output

    HM	17.9.2007	rev 1.2
    	replaced time() with T_PLC_MS() for compatibility reasons
    *)

END_FUNCTION_BLOCK

(* ---- SH_2.st ---- *)
FUNCTION_BLOCK SH_2
    (*http://www.oscat.de/images/OSCATBasic/oscat_basic333_en.pdf#page=301*)
    (* read system time *)
    tx := UDINT_TO_TIME(T_PLC_MS());
    d2 := SHR(DISC,1);

    IF tx - last >= PT THEN
    	last := tx;
    	TRIG := TRUE;

    	(* limit M to 0..16 *)
    	M := LIMIT(1,N,16);

    	(* edge detected lets take the sample *)
    	FOR i := M - 1 TO 1 BY -1 DO buf2[i] := buf2[i-1]; END_FOR
    	buf2[0] := IN;
    	OUT := IN;
    	buf := buf2;

    	(* sort the ARRAY lowest value AT 0 *)
    	FOR start := 0 TO M - 2 DO
    		FOR i := start+1 TO M - 1 DO
    			IF buf[start] > buf[i] THEN
    				temp := buf[start];
    				buf[start] := buf[i];
    				buf[i] := temp;
    			END_IF
    		END_FOR
    	END_FOR

    	(* any calculation with the samples is here *)
    	stop := M - 1 - d2;
    	start := d2;
    	IF NOT EVEN(DISC) THEN start := start + 1; END_IF
    	AVG := 0;
    	FOR i := start TO stop DO AVG := AVG + buf[i]; END_FOR
    	AVG := AVG / INT_TO_REAL(stop - start +1);
    	LOW := buf[start];
    	HIGH := buf[stop];
    ELSE
    	TRIG := FALSE;
    END_IF

    (* revision history
    hm 20. jan. 2007	rev 1.1
    	added input N to specify the amout of samples for average and HIGH LOW calculations
    	added TRIG output

    hm 10. sep. 2007 	rev 1.2
    	an error would be generated if N was set to 0, now N is forced to1 if set to 0.
    	index was OUT of array.

    hm	17. sep. 2007	rev 1.3
    	replaced time() with t_plc_ms() for compatibility reasons

    hm	6. jan. 2008	rev 1.4
    	improved performance

    hm	14. jun. 2008	rev 1.5
    	set default for input N = 16

    hm	10. mar. 2009	rev 1.6
    	added type conversion for compatibility reasons

    *)
END_FUNCTION_BLOCK

(* ---- SH_T.st ---- *)
FUNCTION_BLOCK SH_T
    (*http://www.oscat.de/images/OSCATBasic/oscat_basic333_en.pdf#page=303*)
    IF E THEN OUT := IN; END_IF

    (* revision history
    hm	1. sep. 2006	rev 1.0
    	original version

    hm	18. oct. 2008	rev 1.1
    	changed input en to E for compatibility reasons

    *)
END_FUNCTION_BLOCK

(* ---- SHR_4E.st ---- *)
FUNCTION_BLOCK SHR_4E
    (*http://www.oscat.de/images/OSCATBasic/oscat_basic333_en.pdf#page=249*)
    (* trig.Q signals a rising edge on CLK *)
    trig(CLK := CLK);

    IF SET OR RST THEN
    	Q0 := NOT RST;
    	Q1 := Q0;
    	Q2 := Q0;
    	Q3 := Q0;
    ELSIF trig.Q THEN
    	Q3 := Q2;
    	Q2 := Q1;
    	Q1 := Q0;
    	Q0 := D0;
    END_IF

    (* revision history
    hm	4. aug. 2006	rev 1.0
    	original version

    hm	25. oct. 2008	rev 1.1
    	optimized code

    *)
END_FUNCTION_BLOCK

(* ---- SHR_4UDE.st ---- *)
FUNCTION_BLOCK SHR_4UDE
    (*http://www.oscat.de/images/OSCATBasic/oscat_basic333_en.pdf#page=250*)
    (* trig.Q signals a rising edge on CLK *)
    trig(CLK := CLK);

    IF SET OR RST THEN
    	Q0 := NOT RST;
    	Q1 := Q0;
    	Q2 := Q0;
    	Q3 := Q0;
    ELSIF trig.Q THEN
    	IF DN THEN
    		Q0 := Q1;
    		Q1 := Q2;
    		Q2 := Q3;
    		Q3 := D3;
    	ELSE
    		Q3 := Q2;
    		Q2 := Q1;
    		Q1 := Q0;
    		Q0 := D0;
    	END_IF
    END_IF

    (* revision history
    hm	4. aug. 2006	rev 1.0
    	original version

    hm	25. oct. 2008	rev 1.1
    	optimized code

    hm	14. mar. 2009	rev 1.2
    	removed double assignments

    *)
END_FUNCTION_BLOCK

(* ---- SHR_8PLE.st ---- *)
FUNCTION_BLOCK SHR_8PLE
    (*http://www.oscat.de/images/OSCATBasic/oscat_basic333_en.pdf#page=251*)
    (* flankenerkennung CLK wird high und edge_ war high reset ist nicht aktiv und set ist nicht aktiv *)
    IF CLK AND edge_ AND NOT RST THEN
    	edge_ := FALSE;	(* flanke wurde erkannt und weitere flankenerkennung wird verhindert bis edge_ wieder true ist *)
    	(* hier ist der code für das flankenevent *)
    	IF UP THEN						(*shift UP *)
    		register := SHL(register,1);
    		register.0 := DIN;
    		DOUT := register.7;
    	ELSE								(* shift down *);
    		register := SHR(register,1);
    		register.7 := DIN;
    		DOUT := register.0;
    	END_IF
    	IF LOAD THEN							(* the byte on DIN will be loaded if LOAD = true *)
    		register := DLOAD;
    		IF UP THEN DOUT := register.7; ELSE DOUT := register.0; END_IF
    	END_IF
    END_IF
    IF NOT CLK THEN edge_ := TRUE; END_IF	(* sobald CLK wieder low wird warten auf nächste flanke *)
    IF RST THEN									(* wenn reset aktiv dann ausgang rücksetzen *)
    	register := 0;
    	DOUT := FALSE;
    END_IF

END_FUNCTION_BLOCK

(* ---- SHR_8UDE.st ---- *)
FUNCTION_BLOCK SHR_8UDE
    (*http://www.oscat.de/images/OSCATBasic/oscat_basic333_en.pdf#page=252*)
    (* trig.Q signals a rising edge on CLK *)
    trig(CLK := CLK);

    IF SET OR RST THEN
    	Q0 := NOT RST;
    	Q1 := Q0;
    	Q2 := Q0;
    	Q3 := Q0;
    	Q4 := Q0;
    	Q5 := Q0;
    	Q6 := Q0;
    	Q7 := Q0;
    ELSIF trig.Q THEN
    	IF DN THEN
    		Q0 := Q1;
    		Q1 := Q2;
    		Q2 := Q3;
    		Q3 := Q4;
    		Q4 := Q5;
    		Q5 := Q6;
    		Q6 := Q7;
    		Q7 := D7;
    	ELSE
    		Q7 := Q6;
    		Q6 := Q5;
    		Q5 := Q4;
    		Q4 := Q3;
    		Q3 := Q2;
    		Q2 := Q1;
    		Q1 := Q0;
    		Q0 := D0;
    	END_IF
    END_IF

    (* revision history
    hm	4. aug. 2006	rev 1.0
    	original version

    hm	25. oct. 2008	rev 1.1
    	optimized code

    hm	14. mar. 2009	rev 1.2
    	removed double assignments

    *)
END_FUNCTION_BLOCK

(* ---- SIGNAL.st ---- *)
FUNCTION_BLOCK SIGNAL
    (*http://www.oscat.de/images/OSCATBasic/oscat_basic333_en.pdf#page=468*)
    IF IN THEN
    	(* an alarm is present read system time first *)
    	tx := T_PLC_MS();
    	(* calculate the step counter which is the lowest 3 bits of (time / TS) *)
    	IF TS > t#0s THEN
    		step := UDINT_TO_BYTE(tx / TIME_TO_UDINT(TS) AND 16#0000_0007);
    	ELSE
    		step := UDINT_TO_BYTE(SHR(tx,7) AND 16#0000_0007);
    	END_IF
    	(* convert the value 0-7 IN step into one bit only (bit 0-7) *)
    	step := SHL(one,step);
    	(* generate the output signal *)
    	Q := (step AND SIG) > 0;
    ELSE
    	Q := FALSE;
    END_IF

    (* revision history
    hm	13.12.2007		rev 1.0
    	original version

    *)
END_FUNCTION_BLOCK

(* ---- SIGNAL_4.st ---- *)
FUNCTION_BLOCK SIGNAL_4
    (*http://www.oscat.de/images/OSCATBasic/oscat_basic333_en.pdf#page=469*)
    (* an alarm is present read system time first *)
    (* check if an alarm is present if yes set sig to the alarm pattern otherwise exit the routine *)
    IF IN1 THEN
    	sig(IN := TRUE, SIG := S1, TS := TS);
    ELSIF IN2 THEN
    	sig(IN := TRUE, SIG := S2, TS := TS);
    ELSIF IN3 THEN
    	sig(IN := TRUE, SIG := S3, TS := TS);
    ELSIF IN4 THEN
    	sig(IN := TRUE, SIG := S4, TS := TS);
    ELSE
    	sig(IN := FALSE);
    END_IF

    (* set the output *)
    Q := sig.Q;

    (* revision history
    hm	13.12.2007		rev 1.0
    	original version

    *)

END_FUNCTION_BLOCK

(* ---- SPEED.st ---- *)
FUNCTION_BLOCK SPEED
    (*http://www.oscat.de/images/OSCATBasic/oscat_basic333_en.pdf#page=372*)
    YMS := MS +
    		KMH * 0.27777777777778 +
    		KN * 0.5144444 +
    		MH * 0.44704;
    YKMH := YMS * 3.6;
    YKN := YMS * 1.94384466037535;
    YMH := YMS * 2.23693629205440;

    (*
    Geschwindigkeit Meter durch Sekunde m/s 1 m/s = 3,6 km/h
    km durch (pro) Stunde, nicht „Stundenkilometer“ verwenden
    Knoten KN 1 KN = 1 sm/h = 0,5144 m/s

    *)

    (* revision history
    hm	27. mar. 2009	rev 1.0
    	original version

    hm	11. mar. 2009	rev 1.1
    	improved code

    *)
END_FUNCTION_BLOCK

(* ---- SRAMP.st ---- *)
FUNCTION_BLOCK SRAMP
    (*http://www.oscat.de/images/OSCATBasic/oscat_basic333_en.pdf#page=470*)
    (* read the system_time in microseconds *)
    cycle_time();

    (* assure range of inputs *)
    A_UP := MAX(0.0, A_UP);
    A_DN := MIN(0.0, A_DN);
    VU_MAX := MAX(0.0, VU_MAX);
    VD_MAX := MIN(0.0, VD_MAX);

    (* calculate the output offset *)
    IF RST OR NOT init THEN
    	init := TRUE;
    	Y := 0.0;
    	V := 0.0;
    ELSIF X = Y THEN
    	V := 0.0;
    ELSIF X > Y THEN
    	(* output is too low >> ramp up and brake at the end *)
    	(* accelerate the speed and limit to VU_MAX *)
    	V := MIN(V + A_UP * cycle_time.TC, VU_MAX);
    	(* calculate the max speed to be able to brake and select the lowest *)
    	V := MIN(SQRT((Y-X) * 2.0 * A_DN), V);
    	(* calculate the output and obey limits *)
    	Y := LIMIT(LIMIT_LOW, Y + MIN(V * cycle_time.TC, X-Y), LIMIT_HIGH);
    ELSIF X < Y THEN
    	(* output is too high >> ramp dn and brake at the end *)
    	(* accelerate the speed and limit to VD_MAX *)
    	V := MAX(V + A_DN * cycle_time.TC, VD_MAX);
    	(* calculate the max speed to be able to brake and select the lowest *)
    	V := MAX(-SQRT((Y-X) * 2.0 * A_UP), V);
    	(* calculate the output and obey limits *)
    	Y := LIMIT(LIMIT_LOW, Y + MAX(V * cycle_time.TC, X-Y), LIMIT_HIGH);
    END_IF

    (* revision history
    hm	13. mar. 2008	rev 1.0
    	original version

    hm	11. mar. 2009	rev 1.1
    	real constants updated to new systax using dot

    *)

END_FUNCTION_BLOCK

(* ---- STACK_16.st ---- *)
FUNCTION_BLOCK STACK_16
    (*http://www.oscat.de/images/OSCATBasic/oscat_basic333_en.pdf#page=185*)
    IF RST THEN
    	(* asynchronous reset for the fifo *)
    	pt := 0;
    	EMPTY := TRUE;
    	FULL := FALSE;
    	DOUT := 0;
    ELSIF E THEN
    	IF NOT EMPTY AND RD THEN
    		(* read one element *)
    		pt := pt - 1;
    		DOUT := stack[pt];
    		EMPTY := pt = 0;
    		FULL := FALSE;
    	END_IF
    	IF NOT FULL AND WD THEN
    		(* write one element *)
    		stack[pt] := DIN;
    		pt := pt + 1;
    		FULL := pt > n;
    		EMPTY := FALSE;
    	END_IF
    END_IF

    (* revision history
    hm	4. aug. 2006	rev 1.0
    	original version

    hm	19. feb 2008	rev 1.1
    	performance improvements

    hm	17. oct. 2008	rev 1.2
    	deleted unnecessary init with 0

    hm	27. oct. 2008	rev 1.3
    	optimized performance

    hm	25. jul 2009	rev 2.0
    	changed inputs to allow simultsaneous read and write
    *)

END_FUNCTION_BLOCK

(* ---- STACK_32.st ---- *)
FUNCTION_BLOCK STACK_32
    (*http://www.oscat.de/images/OSCATBasic/oscat_basic333_en.pdf#page=186*)
    IF RST THEN
    	(* asynchronous reset for the fifo *)
    	pt := 0;
    	EMPTY := TRUE;
    	FULL := FALSE;
    	DOUT := 0;
    ELSIF E THEN
    	IF NOT EMPTY AND RD THEN
    		(* read one element *)
    		pt := pt - 1;
    		DOUT := stack[pt];
    		EMPTY := pt = 0;
    		FULL := FALSE;
    	END_IF
    	IF NOT FULL AND WD THEN
    		(* write one element *)
    		stack[pt] := DIN;
    		pt := pt + 1;
    		FULL := pt > n;
    		EMPTY := FALSE;
    	END_IF
    END_IF

    (* revision history
    hm	4. aug. 2006	rev 1.0
    	original version

    hm	19. feb 2008	rev 1.1
    	performance improvements

    hm	17. oct. 2008	rev 1.2
    	deleted unnecessary init with 0

    ks	27. oct. 2008	rev 1.3
    	optimized performance

    hm	25. jul 2009	rev 2.0
    	changed inputs to allow simultsaneous read and write

    *)

END_FUNCTION_BLOCK

(* ---- STAIR2.st ---- *)
FUNCTION_BLOCK STAIR2
    (*http://www.oscat.de/images/OSCATBasic/oscat_basic333_en.pdf#page=304*)
    IF D > 0.0 THEN
    	IF X >= Y + D OR X <= Y - D THEN Y := FLOOR(X/D) * D; END_IF
    ELSE
    	Y := X;
    END_IF

    (* revision history
    hm	28 jan 2007		rev 1.0
    	original version

    hm	27. dec 2007	rev 1.1
    	changed code for better performance

    hm	30. jun. 2008	rev 1.2
    	added type conversions to avoid warnings under codesys 3.0

    ks	26. oct. 2008	rev 1.3
    	improved code

    hm	10. mar. 2009	rev 1.4
    	real constants updated to new systax using dot

    *)
END_FUNCTION_BLOCK
